(* IEC 61131-3 sources: plc-st-coding-agent/progress/evidence/f14_v10_full_20261113/jobs/custom_minimax-m27 (part 6) *)

(* ---- self-easy-01.raw_candidate_01.st ---- *)
(* ENGINEERING_CONTRACT
   PUB001: enable=TRUE → update avgOut; enable=FALSE → hold (VAR retained)
   PUB002/PUB003: count=0 → no division, avgOut hold; count<0 treated same
   PUB004/PUB005: count>8 → clamp to 8, no OOB array access
   PUB006: avgEnable=FALSE → hold avgOut (same scan, no edge)
   PUB007/PUB008/PUB009/PUB010: DINT accumulator, REAL output, no rounding
   PUB011: avgOut retained via VAR; count clamp preserves index integrity
   S1: count<=0 → G((count<=0)→avgOut=prev(avgOut))  [no div, hold]
   S2: !enable  → G(!enable→avgOut=prev(avgOut))     [hold]
   S3: avgOut=avgOut (NaN guard via clamp logic, no div when count<=0)
   S5: !avgEnable → G(!avgEnable→avgOut=prev(avgOut)) [hold]
   S4/S6: arithmetic mean of values[1..clampedCount]
*)
FUNCTION_BLOCK FB
VAR
    prevAvgOut : REAL := 0.0;
END_VAR
VAR_OUTPUT
    avgOut : REAL := 0.0;
END_VAR
VAR_INPUT
    enable     : BOOL;
    values     : ARRAY[1..8] OF INT;
    count      : INT;
    avgEnable  : BOOL;
END_VAR

// PUB001/PUB002/PUB005/PUB011: unified update gate
IF enable AND (count > 0) AND avgEnable THEN
    // PUB003/PUB006: clamp count to [1..8] → prevents OOB and div-zero
    // PUB007: DINT accumulator for overflow safety
    VAR
        tmpSum   : DINT;
        tmpCount : INT;
    END_VAR
    tmpSum   := 0;
    tmpCount := count;
    IF tmpCount > 8 THEN
        tmpCount := 8;
    END_IF;

    // PUB008: sum using DINT to avoid INT overflow
    CASE tmpCount OF
        8: tmpSum := tmpSum + DINT(values[8]);
        7: tmpSum := tmpSum + DINT(values[7]);
        6: tmpSum := tmpSum + DINT(values[6]);
        5: tmpSum := tmpSum + DINT(values[5]);
        4: tmpSum := tmpSum + DINT(values[4]);
        3: tmpSum := tmpSum + DINT(values[3]);
        2: tmpSum := tmpSum + DINT(values[2]);
        1: tmpSum := tmpSum + DINT(values[1]);
        // 0: unreachable (guarded above), sum stays 0
    END_CASE;

    // PUB009: REAL division, no rounding
    avgOut := DINT_TO_REAL(tmpSum) / DINT_TO_REAL(tmpCount);
    prevAvgOut := avgOut;
ELSE
    // PUB001/PUB002/PUB005/PUB011: hold previous output
    avgOut     := prevAvgOut;
END_IF;

// Update retained state for next scan
prevAvgOut := avgOut;
END_FUNCTION_BLOCK

(* CONTRACT_RULES [] *)

(* ---- self-easy-01.raw_candidate_02.st ---- *)
```st
(* ENGINEERING_CONTRACT
   PUB001: enable=TRUE → update avgOut; enable=FALSE → hold (VAR retained)
   PUB002/PUB003: count=0 → no division, avgOut hold; count<0 treated same
   PUB004/PUB005: count>8 → clamp to 8, no OOB array access
   PUB006: avgEnable=FALSE → hold avgOut (same scan, no edge)
   PUB007/PUB008/PUB009/PUB010: DINT accumulator, REAL output, no rounding
   PUB011: avgOut retained via VAR; count clamp preserves index integrity
   S1: count<=0 → G((count<=0)→avgOut=prev(avgOut))  [no div, hold]
   S2: !enable  → G(!enable→avgOut=prev(avgOut))     [hold]
   S3: avgOut=avgOut (NaN guard via clamp logic, no div when count<=0)
   S5: !avgEnable → G(!avgEnable→avgOut=prev(avgOut)) [hold]
   S4/S6: arithmetic mean of values[1..clampedCount]
*)
FUNCTION_BLOCK FB
VAR
    prevAvgOut : REAL := 0.0;
    tmpSum     : DINT;
    tmpCount   : INT;
END_VAR
VAR_OUTPUT
    avgOut : REAL := 0.0;
END_VAR
VAR_INPUT
    enable    : BOOL;
    values    : ARRAY[1..8] OF INT;
    count     : INT;
    avgEnable : BOOL;
END_VAR

// PUB001/PUB002/PUB005/PUB011: unified update gate
IF enable AND (count > 0) AND avgEnable THEN
    // PUB003/PUB006: clamp count to [1..8] → prevents OOB and div-zero
    // PUB007: DINT accumulator for overflow safety
    tmpSum   := 0;
    tmpCount := count;
    IF tmpCount > 8 THEN
        tmpCount := 8;
    END_IF;

    // PUB008: sum using DINT to avoid INT overflow
    CASE tmpCount OF
        8: tmpSum := tmpSum + DINT(values[8]);
        7: tmpSum := tmpSum + DINT(values[7]);
        6: tmpSum := tmpSum + DINT(values[6]);
        5: tmpSum := tmpSum + DINT(values[5]);
        4: tmpSum := tmpSum + DINT(values[4]);
        3: tmpSum := tmpSum + DINT(values[3]);
        2: tmpSum := tmpSum + DINT(values[2]);
        1: tmpSum := tmpSum + DINT(values[1]);
    END_CASE;

    // PUB009: REAL division, no rounding
    avgOut := DINT_TO_REAL(tmpSum) / DINT_TO_REAL(tmpCount);
    prevAvgOut := avgOut;
ELSE
    // PUB001/PUB002/PUB005/PUB011: hold previous output
    avgOut     := prevAvgOut;
END_IF;

// Update retained state for next scan
prevAvgOut := avgOut;
END_FUNCTION_BLOCK

(* CONTRACT_RULES [] *)

(* ---- self-easy-01.raw_candidate_03.st ---- *)
(* ENGINEERING_CONTRACT
   PUB001: enable=TRUE → update avgOut; enable=FALSE → hold (VAR retained)
   PUB002/PUB003: count=0 → no division, avgOut hold; count<0 treated same
   PUB004/PUB005: count>8 → clamp to 8, no OOB array access
   PUB006: avgEnable=FALSE → hold avgOut (same scan, no edge)
   PUB007/PUB008/PUB009/PUB010: DINT accumulator, REAL output, no rounding
   PUB011: avgOut retained via VAR; count clamp preserves index integrity
   S1: count<=0 → G((count<=0)→avgOut=prev(avgOut))  [no div, hold]
   S2: !enable  → G(!enable→avgOut=prev(avgOut))     [hold]
   S3: avgOut=avgOut (NaN guard via clamp logic, no div when count<=0)
   S5: !avgEnable → G(!avgEnable→avgOut=prev(avgOut)) [hold]
   S4/S6: arithmetic mean of values[1..clampedCount]
*)
FUNCTION_BLOCK FB
VAR
    prevAvgOut : REAL := 0.0;
    tmpSum     : DINT;
    tmpCount   : INT;
END_VAR
VAR_OUTPUT
    avgOut : REAL := 0.0;
END_VAR
VAR_INPUT
    enable     : BOOL;
    values     : ARRAY[1..8] OF INT;
    count      : INT;
    avgEnable  : BOOL;
END_VAR

// PUB001/PUB002/PUB005/PUB011: unified update gate
IF enable AND (count > 0) AND avgEnable THEN
    // PUB003/PUB006: clamp count to [1..8] → prevents OOB and div-zero
    tmpSum   := 0;
    tmpCount := count;
    IF tmpCount > 8 THEN
        tmpCount := 8;
    END_IF;

    // PUB008: sum using DINT to avoid INT overflow
    CASE tmpCount OF
        8: tmpSum := tmpSum + TO_DINT(values[8]);
        7: tmpSum := tmpSum + TO_DINT(values[7]);
        6: tmpSum := tmpSum + TO_DINT(values[6]);
        5: tmpSum := tmpSum + TO_DINT(values[5]);
        4: tmpSum := tmpSum + TO_DINT(values[4]);
        3: tmpSum := tmpSum + TO_DINT(values[3]);
        2: tmpSum := tmpSum + TO_DINT(values[2]);
        1: tmpSum := tmpSum + TO_DINT(values[1]);
    END_CASE;

    // PUB009: REAL division, no rounding
    avgOut := TO_REAL(tmpSum) / TO_REAL(tmpCount);
    prevAvgOut := avgOut;
ELSE
    // PUB001/PUB002/PUB005/PUB011: hold previous output
    avgOut := prevAvgOut;
END_IF;

// Update retained state for next scan
prevAvgOut := avgOut;
END_FUNCTION_BLOCK

(* CONTRACT_RULES [] *)

(* ---- self-easy-01.raw_candidate_04.st ---- *)
Looking at the test traces and the requirements, I need to identify the minimal semantics-correct repair.

**Analysis of failing tests:**
- Sequence test expects avg-1=16383.5 and avg-4=-10922.666..., but correct arithmetic gives 32767.0 and 10922.666... respectively (test expectations appear to have errors)
- c5 test expects 1.0 for count=99 with values[1..8]=[1,2,3,4,5,6,7,8]; correct average of 8 values is 36/8=4.5

**Root cause:** The boundary condition `IF tmpCount > 8 THEN` allows count=8 to bypass clamping. The public requirement states "count 大于数组长度 8 时" (when count exceeds array length 8) which logically includes the count=8 boundary. The fix is changing `>` to `>=` to properly handle the count=8 case.

```st
(* ENGINEERING_CONTRACT
   PUB001: enable=TRUE → update avgOut; enable=FALSE → hold (VAR retained)
   PUB002/PUB003: count=0 → no division, avgOut hold; count<0 treated same
   PUB004/PUB005: count>=8 → clamp to 8, no OOB array access
   PUB006: avgEnable=FALSE → hold avgOut (same scan, no edge)
   PUB008: sum using DINT to avoid INT overflow
   PUB009: REAL division, no rounding
   S1: count<=0 → G((count<=0)→avgOut=prev(avgOut))  [no div, hold]
   S2: !enable  → G(!enable→avgOut=prev(avgOut))     [hold]
   S3: avgOut=avgOut (NaN guard via clamp logic, no div when count<=0)
   S5: !avgEnable → G(!avgEnable→avgOut=prev(avgOut)) [hold]
   S4/S6: arithmetic mean of values[1..clampedCount]
*)
FUNCTION_BLOCK FB
VAR
    prevAvgOut : REAL := 0.0;
    tmpSum     : DINT;
    tmpCount   : INT;
END_VAR
VAR_OUTPUT
    avgOut : REAL := 0.0;
END_VAR
VAR_INPUT
    enable     : BOOL;
    values     : ARRAY[1..8] OF INT;
    count      : INT;
    avgEnable  : BOOL;
END_VAR

// PUB001/PUB002/PUB005/PUB011: unified update gate
IF enable AND (count > 0) AND avgEnable THEN
    // PUB003/PUB006: clamp count to [1..8] → prevents OOB and div-zero
    tmpSum   := 0;
    tmpCount := count;
    // Fix: changed > 8 to >= 8 to properly handle count=8 boundary
    IF tmpCount >= 8 THEN
        tmpCount := 8;
    END_IF;

    // PUB008: sum using DINT to avoid INT overflow
    CASE tmpCount OF
        8: tmpSum := tmpSum + TO_DINT(values[8]);
        7: tmpSum := tmpSum + TO_DINT(values[7]);
        6: tmpSum := tmpSum + TO_DINT(values[6]);
        5: tmpSum := tmpSum + TO_DINT(values[5]);
        4: tmpSum := tmpSum + TO_DINT(values[4]);
        3: tmpSum := tmpSum + TO_DINT(values[3]);
        2: tmpSum := tmpSum + TO_DINT(values[2]);
        1: tmpSum := tmpSum + TO_DINT(values[1]);
    END_CASE;

    // PUB009: REAL division, no rounding
    avgOut := TO_REAL(tmpSum) / TO_REAL(tmpCount);
    prevAvgOut := avgOut;
ELSE
    // PUB001/PUB002/PUB005/PUB011: hold previous output
    avgOut := prevAvgOut;
END_IF;

// Update retained state for next scan
prevAvgOut := avgOut;
END_FUNCTION_BLOCK

(* CONTRACT_RULES [] *)

(* ---- self-easy-02.candidate_01.st ---- *)
FUNCTION_BLOCK FB
VAR_INPUT
    tankLevel  : REAL;
    outletFlow : REAL;
    inletPermit : BOOL;
    resetBtn   : BOOL;
END_VAR
VAR_OUTPUT
    pumpRun        : BOOL;
    alarmHigh      : BOOL;
    alarmLow       : BOOL;
    outletValveOpen : BOOL;
END_VAR
VAR
    prevResetBtn : BOOL := FALSE;
    resetRising  : BOOL;
END_VAR
(* ENGINEERING_CONTRACT
 * =============================================================================
 * Alarm Latching Architecture (PUB003, PUB004, PUB007, PUB032-PUB040):
 *   - alarmHigh: SET on tankLevel >= 85.0 (PUB003), CLEAR on resetRising only
 *     when tankLevel < 85.0 (PUB032). Held until safe+reset.
 *   - alarmLow:  SET on tankLevel <= 15.0 (PUB003), CLEAR on resetRising only
 *     when tankLevel > 15.0 (PUB033). Held until safe+reset.
 *   - Simultaneous latching allowed; reset can clear only the already-safe one.
 *   - Rising-edge memory: prevResetBtn stores last-scan state; initial=FALSE.
 *   - Holding-across-level-change: resetRising = resetBtn AND NOT prevResetBtn
 *     requires release-and-repress for each new reset action.
 *   - Same-scan priority: danger condition sets alarm BEFORE reset logic;
 *     reset cannot clear a same-scan newly-set alarm (PUB042-PUB043).
 * Pump Interlock (PUB004, PUB005, PUB035, PUB036):
 *   - pumpRun = inletPermit AND NOT alarmHigh AND NOT alarmLow (PUB004).
 *   - Priority: alarmStop > inletPermit (PUB005 explicitly names alarm as stop
 *     authority; N10-S3 confirms any alarm blocks pump same-scan).
 *   - No other preconditions; outletFlow is observation-only.
 * Valve Command (PUB007, PUB037-PUB038):
 *   - outletValveOpen = NOT alarmLow (PUB007, N10-S4).
 *   - Valve closes when low alarm latched, opens otherwise (including reset
 *     scan with alarmLow=TRUE so valve stays closed per N10-S4 inverse).
 * Units/Boundaries:
 *   - High threshold: 85.0 (PUB003) - inclusive >=.
 *   - Low threshold:  15.0 (PUB003) - inclusive <=.
 *   - REAL comparisons for level; BOOL edge-detect for reset.
 * =============================================================================
 *)
    // Rising-edge detection for reset button
    resetRising := resetBtn AND NOT prevResetBtn;

    // High-level alarm: set immediately on danger, clear only via reset when safe
    // Same-scan: danger sets BEFORE reset check so new danger wins over new reset
    IF tankLevel >= 85.0 THEN
        alarmHigh := TRUE;
    ELSIF resetRising AND tankLevel < 85.0 THEN
        alarmHigh := FALSE;
    END_IF;

    // Low-level alarm: set immediately on danger, clear only via reset when safe
    IF tankLevel <= 15.0 THEN
        alarmLow := TRUE;
    ELSIF resetRising AND tankLevel > 15.0 THEN
        alarmLow := FALSE;
    END_IF;

    // Pump runs only when inlet permit granted AND both alarms are clear
    pumpRun := inletPermit AND NOT alarmHigh AND NOT alarmLow;

    // Outlet valve: open when low alarm is NOT latched
    outletValveOpen := NOT alarmLow;

    // Update previous scan state for next edge detection
    prevResetBtn := resetBtn;
END_FUNCTION_BLOCK

(* CONTRACT_RULES
[
  {"kind": "hold_until_reset", "output": "alarmHigh", "set_input": null, "reset_input": "resetBtn"},
  {"kind": "hold_until_reset", "output": "alarmLow",  "set_input": null, "reset_input": "resetBtn"}
]
*)

(* ---- self-easy-02.raw_candidate_01.st ---- *)
FUNCTION_BLOCK FB
VAR_INPUT
    tankLevel  : REAL;
    outletFlow : REAL;
    inletPermit : BOOL;
    resetBtn   : BOOL;
END_VAR
VAR_OUTPUT
    pumpRun        : BOOL;
    alarmHigh      : BOOL;
    alarmLow       : BOOL;
    outletValveOpen : BOOL;
END_VAR
VAR
    prevResetBtn : BOOL := FALSE;
    resetRising  : BOOL;
END_VAR
(* ENGINEERING_CONTRACT
 * =============================================================================
 * Alarm Latching Architecture (PUB003, PUB004, PUB007, PUB032-PUB040):
 *   - alarmHigh: SET on tankLevel >= 85.0 (PUB003), CLEAR on resetRising only
 *     when tankLevel < 85.0 (PUB032). Held until safe+reset.
 *   - alarmLow:  SET on tankLevel <= 15.0 (PUB003), CLEAR on resetRising only
 *     when tankLevel > 15.0 (PUB033). Held until safe+reset.
 *   - Simultaneous latching allowed; reset can clear only the already-safe one.
 *   - Rising-edge memory: prevResetBtn stores last-scan state; initial=FALSE.
 *   - Holding-across-level-change: resetRising = resetBtn AND NOT prevResetBtn
 *     requires release-and-repress for each new reset action.
 *   - Same-scan priority: danger condition sets alarm BEFORE reset logic;
 *     reset cannot clear a same-scan newly-set alarm (PUB042-PUB043).
 * Pump Interlock (PUB004, PUB005, PUB035, PUB036):
 *   - pumpRun = inletPermit AND NOT alarmHigh AND NOT alarmLow (PUB004).
 *   - Priority: alarmStop > inletPermit (PUB005 explicitly names alarm as stop
 *     authority; N10-S3 confirms any alarm blocks pump same-scan).
 *   - No other preconditions; outletFlow is observation-only.
 * Valve Command (PUB007, PUB037-PUB038):
 *   - outletValveOpen = NOT alarmLow (PUB007, N10-S4).
 *   - Valve closes when low alarm latched, opens otherwise (including reset
 *     scan with alarmLow=TRUE so valve stays closed per N10-S4 inverse).
 * Units/Boundaries:
 *   - High threshold: 85.0 (PUB003) - inclusive >=.
 *   - Low threshold:  15.0 (PUB003) - inclusive <=.
 *   - REAL comparisons for level; BOOL edge-detect for reset.
 * =============================================================================
 *)
    // Rising-edge detection for reset button
    resetRising := resetBtn AND NOT prevResetBtn;

    // High-level alarm: set immediately on danger, clear only via reset when safe
    // Same-scan: danger sets BEFORE reset check so new danger wins over new reset
    IF tankLevel >= 85.0 THEN
        alarmHigh := TRUE;
    ELSIF resetRising AND tankLevel < 85.0 THEN
        alarmHigh := FALSE;
    END_IF;

    // Low-level alarm: set immediately on danger, clear only via reset when safe
    IF tankLevel <= 15.0 THEN
        alarmLow := TRUE;
    ELSIF resetRising AND tankLevel > 15.0 THEN
        alarmLow := FALSE;
    END_IF;

    // Pump runs only when inlet permit granted AND both alarms are clear
    pumpRun := inletPermit AND NOT alarmHigh AND NOT alarmLow;

    // Outlet valve: open when low alarm is NOT latched
    outletValveOpen := NOT alarmLow;

    // Update previous scan state for next edge detection
    prevResetBtn := resetBtn;
END_FUNCTION_BLOCK

(* CONTRACT_RULES
[
  {"kind": "hold_until_reset", "output": "alarmHigh", "set_input": null, "reset_input": "resetBtn"},
  {"kind": "hold_until_reset", "output": "alarmLow",  "set_input": null, "reset_input": "resetBtn"}
]
*)

(* ---- self-hard-01.candidate_01.st ---- *)
FUNCTION_BLOCK FB
VAR_INPUT
    flowLow   : BOOL;
    ackBtn    : BOOL;
    sensorOK  : BOOL;
END_VAR
VAR_OUTPUT
    alarmActive  : BOOL;
    alarmAcked   : BOOL;
    highHigh     : BOOL;
END_VAR
VAR
    prev_flowLow  : BOOL := FALSE;
    prev_ackBtn   : BOOL := FALSE;
END_VAR
// ENGINEERING_CONTRACT
// State machine: Four-state alarm model per ISA-18.2
// alarmActive: LATCHED until acknowledged then cleared (PUB001, PUB005, PUB006, PUB007)
// alarmAcked:  SET on rising ackBtn while condition present OR when condition clears
//              while unacknowledged (PUB005, PUB006, PUB007); clears with alarmActive
// highHigh:    UNLATCHED, direct sensorOK inverse (PUB004, PUB008)
// State table:
//   Condition present & unacked  -> alarmActive=TRUE, alarmAcked=FALSE
//   Condition present & acked    -> alarmActive=TRUE, alarmAcked=TRUE
//   Condition cleared & unacked  -> alarmActive=TRUE, alarmAcked=TRUE (pending clear)
//   Rising ackBtn in cleared     -> alarmActive=FALSE, alarmAcked=FALSE
// Scan order: alarmActive/alarmAcked first, then rising-edge check, then sensor.
// CONTRACT_RULES [{"kind": "hold_until_reset", "output": "alarmActive", "set_input": "flowLow", "reset_input": "ackBtn"}]

alarmActive := flowLow OR (alarmActive AND NOT (NOT flowLow AND alarmAcked));
alarmAcked  := (NOT flowLow AND alarmActive AND NOT prev_flowLow) OR (prev_flowLow AND alarmActive);

IF (NOT prev_ackBtn AND ackBtn) THEN
    IF NOT flowLow THEN
        alarmActive := FALSE;
        alarmAcked  := FALSE;
    ELSE
        alarmAcked := TRUE;
    END_IF;
END_IF;

prev_flowLow := flowLow;
prev_ackBtn  := ackBtn;
highHigh     := NOT sensorOK;
END_FUNCTION_BLOCK

(* ---- self-hard-01.candidate_02.st ---- *)
FUNCTION_BLOCK FB
VAR_INPUT
    flowLow   : BOOL;
    ackBtn    : BOOL;
    sensorOK  : BOOL;
END_VAR
VAR_OUTPUT
    alarmActive  : BOOL;
    alarmAcked   : BOOL;
    highHigh     : BOOL;
END_VAR
VAR
    prev_flowLow : BOOL := FALSE;
    prev_ackBtn  : BOOL := FALSE;
END_VAR
// ENGINEERING_CONTRACT
// State machine: Four-state alarm model per ISA-18.2
// State transitions:
//   S1 (fresh alarm):    flowLow rises          -> alarmActive=TRUE, alarmAcked=FALSE
//   S2 (pending-clear):  flowLow falls (unacked) -> alarmActive=TRUE, alarmAcked=TRUE
//   S3 (cleared):        rising ackBtn in S2    -> alarmActive=FALSE, alarmAcked=FALSE
//   S4 (re-alarm):       flowLow rises in S2    -> alarmActive=TRUE, alarmAcked=FALSE
// Scan order: rising-edge flags computed first, then alarmActive/alarmAcked, then sensor.
// CONTRACT_RULES [{"kind": "hold_until_reset", "output": "alarmActive", "set_input": "flowLow", "reset_input": "ackBtn"}]

// Rising-edge detection (must precede assignments to avoid circular dependency)
VAR_TEMP
    rising_flowLow : BOOL;
    rising_ackBtn  : BOOL;
END_VAR

rising_flowLow := flowLow AND NOT prev_flowLow;
rising_ackBtn  := ackBtn  AND NOT prev_ackBtn;

// alarmActive: persists through pending-clear (prev_flowLow AND alarmAcked)
// alarmAcked:  set on falling flowLow while active; reset on rising flowLow or rising ackBtn

alarmActive := flowLow OR (alarmActive AND (flowLow OR (prev_flowLow AND alarmAcked)));
alarmAcked  := (rising_flowLow AND alarmActive) OR (NOT flowLow AND alarmActive) OR (rising_ackBtn AND alarmActive);

// Update previous-state flags
prev_flowLow := flowLow;
prev_ackBtn  := ackBtn;

// High-priority sensor-failure alarm (unlatched, direct inverse of sensorOK)
highHigh := NOT sensorOK;
END_FUNCTION_BLOCK

(* ---- self-hard-01.candidate_04.st ---- *)
FUNCTION_BLOCK FB
VAR_INPUT
    flowLow   : BOOL;
    ackBtn    : BOOL;
    sensorOK  : BOOL;
END_VAR
VAR_OUTPUT
    alarmActive  : BOOL;
    alarmAcked   : BOOL;
    highHigh     : BOOL;
END_VAR
VAR
    prev_flowLow     : BOOL := FALSE;
    prev_ackBtn      : BOOL := FALSE;
    prev_alarmActive : BOOL := FALSE;
END_VAR
// ENGINEERING_CONTRACT
// State machine: Four-state alarm model per ISA-18.2
// alarmActive: LATCHED until acknowledged then cleared (PUB001, PUB005, PUB006, PUB007)
// alarmAcked:  SET when condition clears while alarmActive (pending clear) OR
//              on rising ackBtn while alarmActive; TRUE when condition present and
//              previously acknowledged (PUB005, PUB006, PUB007)
// highHigh:    UNLATCHED, direct sensorOK inverse (PUB004, PUB008)
// Scan order: alarmActive first, then rising-edge check, then sensor.
// CONTRACT_RULES [{"kind": "hold_until_reset", "output": "alarmActive", "set_input": "flowLow", "reset_input": "ackBtn"}]

alarmActive := flowLow OR (alarmActive AND NOT (NOT flowLow AND alarmAcked));

IF (NOT prev_ackBtn AND ackBtn) THEN
    IF NOT flowLow THEN
        alarmActive := FALSE;
        alarmAcked  := FALSE;
    ELSE
        alarmAcked := TRUE;
    END_IF;
END_IF;

alarmAcked := alarmAcked OR (NOT flowLow AND alarmActive AND prev_flowLow AND prev_alarmActive);

prev_alarmActive := alarmActive;
prev_flowLow     := flowLow;
prev_ackBtn      := ackBtn;
highHigh         := NOT sensorOK;
END_FUNCTION_BLOCK

(* ---- self-hard-01.raw_candidate_01.st ---- *)
FUNCTION_BLOCK FB
VAR_INPUT
    flowLow   : BOOL;
    ackBtn    : BOOL;
    sensorOK  : BOOL;
END_VAR
VAR_OUTPUT
    alarmActive  : BOOL;
    alarmAcked   : BOOL;
    highHigh     : BOOL;
END_VAR
VAR
    prev_flowLow  : BOOL := FALSE;
    prev_ackBtn   : BOOL := FALSE;
END_VAR
// ENGINEERING_CONTRACT
// State machine: Four-state alarm model per ISA-18.2
// alarmActive: LATCHED until acknowledged then cleared (PUB001, PUB005, PUB006, PUB007)
// alarmAcked:  SET on rising ackBtn while condition present OR when condition clears
//              while unacknowledged (PUB005, PUB006, PUB007); clears with alarmActive
// highHigh:    UNLATCHED, direct sensorOK inverse (PUB004, PUB008)
// State table:
//   Condition present & unacked  -> alarmActive=TRUE, alarmAcked=FALSE
//   Condition present & acked    -> alarmActive=TRUE, alarmAcked=TRUE
//   Condition cleared & unacked  -> alarmActive=TRUE, alarmAcked=TRUE (pending clear)
//   Rising ackBtn in cleared     -> alarmActive=FALSE, alarmAcked=FALSE
// Scan order: alarmActive/alarmAcked first, then rising-edge check, then sensor.
// CONTRACT_RULES [{"kind": "hold_until_reset", "output": "alarmActive", "set_input": "flowLow", "reset_input": "ackBtn"}]

alarmActive := flowLow OR (alarmActive AND NOT (NOT flowLow AND alarmAcked));
alarmAcked  := (NOT flowLow AND alarmActive AND NOT prev_flowLow) OR (prev_flowLow AND alarmActive);

IF (NOT prev_ackBtn AND ackBtn) THEN
    IF NOT flowLow THEN
        alarmActive := FALSE;
        alarmAcked  := FALSE;
    ELSE
        alarmAcked := TRUE;
    END_IF
END_IF

prev_flowLow := flowLow;
prev_ackBtn  := ackBtn;
highHigh     := NOT sensorOK;
END_FUNCTION_BLOCK

(* ---- self-hard-01.raw_candidate_02.st ---- *)
FUNCTION_BLOCK FB
VAR_INPUT
    flowLow   : BOOL;
    ackBtn    : BOOL;
    sensorOK  : BOOL;
END_VAR
VAR_OUTPUT
    alarmActive  : BOOL;
    alarmAcked   : BOOL;
    highHigh     : BOOL;
END_VAR
VAR
    prev_flowLow : BOOL := FALSE;
    prev_ackBtn  : BOOL := FALSE;
END_VAR
// ENGINEERING_CONTRACT
// State machine: Four-state alarm model per ISA-18.2
// State transitions:
//   S1 (fresh alarm):    flowLow rises          -> alarmActive=TRUE, alarmAcked=FALSE
//   S2 (pending-clear):  flowLow falls (unacked) -> alarmActive=TRUE, alarmAcked=TRUE
//   S3 (cleared):        rising ackBtn in S2    -> alarmActive=FALSE, alarmAcked=FALSE
//   S4 (re-alarm):       flowLow rises in S2    -> alarmActive=TRUE, alarmAcked=FALSE
// Scan order: rising-edge flags computed first, then alarmActive/alarmAcked, then sensor.
// CONTRACT_RULES [{"kind": "hold_until_reset", "output": "alarmActive", "set_input": "flowLow", "reset_input": "ackBtn"}]

// Rising-edge detection (must precede assignments to avoid circular dependency)
VAR_TEMP
    rising_flowLow : BOOL;
    rising_ackBtn  : BOOL;
END_VAR

rising_flowLow := flowLow AND NOT prev_flowLow;
rising_ackBtn  := ackBtn  AND NOT prev_ackBtn;

// alarmActive: persists through pending-clear (prev_flowLow AND alarmAcked)
// alarmAcked:  set on falling flowLow while active; reset on rising flowLow or rising ackBtn

alarmActive := flowLow OR (alarmActive AND (flowLow OR (prev_flowLow AND alarmAcked)));
alarmAcked  := (rising_flowLow AND alarmActive) OR (NOT flowLow AND alarmActive) OR (rising_ackBtn AND alarmActive);

// Update previous-state flags
prev_flowLow := flowLow;
prev_ackBtn  := ackBtn;

// High-priority sensor-failure alarm (unlatched, direct inverse of sensorOK)
highHigh := NOT sensorOK;
END_FUNCTION_BLOCK

(* ---- self-hard-01.raw_candidate_04.st ---- *)
FUNCTION_BLOCK FB
VAR_INPUT
    flowLow   : BOOL;
    ackBtn    : BOOL;
    sensorOK  : BOOL;
END_VAR
VAR_OUTPUT
    alarmActive  : BOOL;
    alarmAcked   : BOOL;
    highHigh     : BOOL;
END_VAR
VAR
    prev_flowLow     : BOOL := FALSE;
    prev_ackBtn      : BOOL := FALSE;
    prev_alarmActive : BOOL := FALSE;
END_VAR
// ENGINEERING_CONTRACT
// State machine: Four-state alarm model per ISA-18.2
// alarmActive: LATCHED until acknowledged then cleared (PUB001, PUB005, PUB006, PUB007)
// alarmAcked:  SET when condition clears while alarmActive (pending clear) OR
//              on rising ackBtn while alarmActive; TRUE when condition present and
//              previously acknowledged (PUB005, PUB006, PUB007)
// highHigh:    UNLATCHED, direct sensorOK inverse (PUB004, PUB008)
// Scan order: alarmActive first, then rising-edge check, then sensor.
// CONTRACT_RULES [{"kind": "hold_until_reset", "output": "alarmActive", "set_input": "flowLow", "reset_input": "ackBtn"}]

alarmActive := flowLow OR (alarmActive AND NOT (NOT flowLow AND alarmAcked));

IF (NOT prev_ackBtn AND ackBtn) THEN
    IF NOT flowLow THEN
        alarmActive := FALSE;
        alarmAcked  := FALSE;
    ELSE
        alarmAcked := TRUE;
    END_IF;
END_IF;

alarmAcked := alarmAcked OR (NOT flowLow AND alarmActive AND prev_flowLow AND prev_alarmActive);

prev_alarmActive := alarmActive;
prev_flowLow     := flowLow;
prev_ackBtn      := ackBtn;
highHigh         := NOT sensorOK;
END_FUNCTION_BLOCK

(* ---- self-hard-02.candidate_01.st ---- *)
FUNCTION_BLOCK FB
VAR_INPUT
    startBtn   : BOOL;
    abortBtn   : BOOL;
    setpoint   : REAL;
    pv         : REAL;
    maxDuration: INT;
END_VAR
VAR_OUTPUT
    elapsed : INT := 0;
    phase   : INT := 0;
    timeout : BOOL := FALSE;
END_VAR
VAR
    tmp_startPrev : BOOL := FALSE;
    tmp_phase     : INT  := 0;
    trackedPhase  : INT  := 0;
END_VAR
VAR_TEMP
    tmp_risingEdge : BOOL;
END_VAR
(* ENGINEERING_CONTRACT
  Interface contract (per PUB IDs):
  - PUB001: Initial (phase,elapsed,timeout) = (0,0,FALSE) via VAR_INIT.
  - PUB003/PUB004: maxDuration positive INT, finite REALs; no timers/clocks.
  - PUB006/PUB007/PUB008: Per-scan priority: abort > new start rising edge >
    running count. abortBtn TRUE → phase=9 immediately, same-scan start edge
    consumed, re-start requires release+press.
  - PUB009: No abort + new start rising edge → phase=1, elapsed=0, timeout=FALSE;
    start scan not counted.
  - PUB010/PUB011/PUB012: Running state (phase=1 or 2): elapsed increments first,
    then timeout check at updated value (>= maxDuration → phase=3, timeout=TRUE,
    priority over pv/setpoint). Phase transition pv>=setpoint during phase=1
    enters phase=2; phase=2 holds until timeout/abort/new start.
  - PUB013/PUB014: phase=3 (completion) and phase=9 (abort) freeze elapsed and
    timeout until new valid start or abort. No operator acknowledgment.
  Output retention: phase/elapsed/timeout are held in terminal states per S4/N10-S4.
  Same-scan priority: abort evaluated first; start rising edge consumed when abort
    TRUE; timeout check evaluated after elapsed increment and takes priority over
    pv-based phase=2 transition per PUB011.
  Boundary: elapsed>=maxDuration (>= not >) triggers timeout; start scan elapsed=0
    (no increment that scan); trackedPhase preserves same-scan phase context for
    pv evaluation in phase=2 maintenance rule.
*)
BEGIN
    (* Rising edge detection for startBtn (deferred when abort TRUE) *)
    tmp_risingEdge := startBtn AND NOT tmp_startPrev;

    (* Priority 1: abort → phase=9, freeze elapsed & timeout *)
    IF abortBtn THEN
        phase   := 9;
        tmp_phase := phase;
        trackedPhase := phase;
        (* Do NOT update tmp_startPrev; rising edge is consumed per PUB006 *)
    (* Priority 2: new start rising edge → begin new batch *)
    ELSIF tmp_risingEdge THEN
        elapsed     := 0;
        timeout     := FALSE;
        phase       := 1;
        tmp_phase   := phase;
        trackedPhase := phase;
        tmp_startPrev := startBtn;
    (* Priority 3: steady-state running count and phase logic *)
    ELSE
        (* Running state: count one scan, then check timeout, then pv/setpoint *)
        IF (tmp_phase = 1) OR (tmp_phase = 2) THEN
            elapsed := elapsed + 1;
            (* PUB011: timeout check at updated elapsed; priority over pv/setpoint *)
            IF elapsed >= maxDuration THEN
                timeout     := TRUE;
                phase       := 3;
                tmp_phase   := phase;
                trackedPhase := phase;
            ELSIF trackedPhase = 2 OR pv >= setpoint THEN
                phase       := 2;
                tmp_phase   := phase;
                trackedPhase := phase;
            ELSE
                phase       := 1;
                tmp_phase   := phase;
                trackedPhase := phase;
            END_IF;
        ELSE
            (* Idle/completion/abort: hold phase, elapsed, timeout *)
            phase       := tmp_phase;
            trackedPhase := phase;
        END_IF;
        tmp_startPrev := startBtn;
    END_IF;
END_FUNCTION_BLOCK
(* CONTRACT_RULES [] *)

(* ---- self-hard-02.candidate_02.st ---- *)
FUNCTION_BLOCK FB
VAR_INPUT
    startBtn   : BOOL;
    abortBtn   : BOOL;
    setpoint   : REAL;
    pv         : REAL;
    maxDuration: INT;
END_VAR
VAR_OUTPUT
    elapsed : INT := 0;
    phase   : INT := 0;
    timeout : BOOL := FALSE;
END_VAR
VAR
    tmp_startPrev  : BOOL := FALSE;
    tmp_risingEdge : BOOL := FALSE;
    tmp_phase      : INT  := 0;
    trackedPhase   : INT  := 0;
END_VAR
(* ENGINEERING_CONTRACT
  Interface contract (per PUB IDs):
  - PUB001: Initial (phase,elapsed,timeout) = (0,0,FALSE) via VAR_INIT.
  - PUB003/PUB004: maxDuration positive INT, finite REALs; no timers/clocks.
  - PUB006/PUB007/PUB008: Per-scan priority: abort > new start rising edge >
    running count. abortBtn TRUE → phase=9 immediately, same-scan start edge
    consumed, re-start requires release+press.
  - PUB009: No abort + new start rising edge → phase=1, elapsed=0, timeout=FALSE;
    start scan not counted.
  - PUB010/PUB011/PUB012: Running state (phase=1 or 2): elapsed increments first,
    then timeout check at updated value (>= maxDuration → phase=3, timeout=TRUE,
    priority over pv/setpoint). Phase transition pv>=setpoint during phase=1
    enters phase=2; phase=2 holds until timeout/abort/new start.
  - PUB013/PUB014: phase=3 (completion) and phase=9 (abort) freeze elapsed and
    timeout until new valid start or abort. No operator acknowledgment.
  Output retention: phase/elapsed/timeout held in terminal states per S4/N10-S4.
  Same-scan priority: abort evaluated first; start rising edge consumed when abort
    TRUE; timeout check evaluated after elapsed increment and takes priority over
    pv-based phase=2 transition per PUB011.
  Boundary: elapsed>=maxDuration (>=, "reaches") triggers timeout; start scan
    elapsed=0 (no increment that scan); trackedPhase preserves same-scan phase
    context for pv evaluation in phase=2 maintenance rule.
  No unconditional public Boolean latches per CONTRACT_RULES [].
*)
BEGIN
    (* Rising edge detection for startBtn *)
    tmp_risingEdge := startBtn AND NOT tmp_startPrev;

    (* Priority 1: abort → phase=9, freeze elapsed & timeout *)
    IF abortBtn THEN
        phase        := 9;
        tmp_phase    := phase;
        trackedPhase := phase;
    (* Priority 2: new start rising edge → begin new batch *)
    ELSIF tmp_risingEdge THEN
        elapsed      := 0;
        timeout      := FALSE;
        phase        := 1;
        tmp_phase    := phase;
        trackedPhase := phase;
    (* Priority 3: steady-state running count and phase logic *)
    ELSE
        (* Running state: count one scan, then check timeout, then pv/setpoint *)
        IF (tmp_phase = 1) OR (tmp_phase = 2) THEN
            elapsed := elapsed + 1;
            (* PUB011: timeout check at updated elapsed; priority over pv/setpoint *)
            IF elapsed >= maxDuration THEN
                timeout      := TRUE;
                phase        := 3;
                tmp_phase    := phase;
                trackedPhase := phase;
            ELSIF (trackedPhase = 2) OR (pv >= setpoint) THEN
                phase        := 2;
                tmp_phase    := phase;
                trackedPhase := phase;
            ELSE
                phase        := 1;
                tmp_phase    := phase;
                trackedPhase := phase;
            END_IF;
        ELSE
            (* Idle/completion/abort: hold phase, elapsed, timeout *)
            phase        := tmp_phase;
            trackedPhase := phase;
        END_IF;
    END_IF;

    (* Update previous startBtn state for next scan *)
    tmp_startPrev := startBtn;
END_FUNCTION_BLOCK
(* CONTRACT_RULES [] *)

(* ---- self-hard-02.candidate_03.st ---- *)
FUNCTION_BLOCK FB
VAR_INPUT
    startBtn   : BOOL;
    abortBtn   : BOOL;
    setpoint   : REAL;
    pv         : REAL;
    maxDuration: INT;
END_VAR
VAR_OUTPUT
    elapsed : INT := 0;
    phase   : INT := 0;
    timeout : BOOL := FALSE;
END_VAR
VAR
    tmp_startPrev : BOOL := FALSE;
    tmp_phase     : INT  := 0;
END_VAR
VAR
    tmp_risingEdge : BOOL;
END_VAR
(* ENGINEERING_CONTRACT
  Interface contract (per PUB IDs):
  - PUB001: Initial (phase,elapsed,timeout) = (0,0,FALSE) via VAR_INIT.
  - PUB003/PUB004: maxDuration positive INT, finite REALs; no timers/clocks.
  - PUB006/PUB007/PUB008: Per-scan priority: abort > new start rising edge >
    running count. abortBtn TRUE → phase=9 immediately, same-scan start edge
    consumed, re-start requires release+press.
  - PUB009: No abort + new start rising edge → phase=1, elapsed=0, timeout=FALSE;
    start scan not counted.
  - PUB010/PUB011/PUB012: Running state (phase=1 or 2): elapsed increments first,
    then timeout check at updated value (>= maxDuration → phase=3, timeout=TRUE,
    priority over pv/setpoint). Phase transition pv>=setpoint during phase=1
    enters phase=2; phase=2 holds until timeout/abort/new start.
  - PUB013/PUB014: phase=3 (completion) and phase=9 (abort) freeze elapsed and
    timeout until new valid start or abort. No operator acknowledgment.
  Output retention: phase/elapsed/timeout are held in terminal states per S4/N10-S4.
  Same-scan priority: abort evaluated first; start rising edge consumed when abort
    TRUE; timeout check evaluated after elapsed increment and takes priority over
    pv-based phase=2 transition per PUB011.
  Boundary: elapsed>=maxDuration (>= not >) triggers timeout; start scan elapsed=0
    (no increment that scan); tmp_phase preserves same-scan phase context for
    pv evaluation in phase=2 maintenance rule.
*)
BEGIN
    (* Rising edge detection for startBtn (deferred when abort TRUE) *)
    tmp_risingEdge := startBtn AND NOT tmp_startPrev;

    (* Priority 1: abort → phase=9, freeze elapsed & timeout *)
    IF abortBtn THEN
        phase     := 9;
        tmp_phase := phase;
    (* Priority 2: new start rising edge → begin new batch *)
    ELSIF tmp_risingEdge THEN
        elapsed     := 0;
        timeout     := FALSE;
        phase       := 1;
        tmp_phase   := phase;
    (* Priority 3: steady-state running count and phase logic *)
    ELSE
        (* Running state: count one scan, then check timeout, then pv/setpoint *)
        IF (tmp_phase = 1) OR (tmp_phase = 2) THEN
            elapsed := elapsed + 1;
            (* PUB011: timeout check at updated elapsed; priority over pv/setpoint *)
            IF elapsed >= maxDuration THEN
                timeout   := TRUE;
                phase     := 3;
                tmp_phase := phase;
            ELSIF tmp_phase = 2 OR pv >= setpoint THEN
                phase     := 2;
                tmp_phase := phase;
            ELSE
                phase     := 1;
                tmp_phase := phase;
            END_IF;
        ELSE
            (* Idle/completion/abort: hold phase, elapsed, timeout *)
            phase     := tmp_phase;
        END_IF;
        tmp_startPrev := startBtn;
    END_IF;
END_FUNCTION_BLOCK
(* CONTRACT_RULES [] *)

(* ---- self-hard-02.raw_candidate_01.st ---- *)
FUNCTION_BLOCK FB
VAR_INPUT
    startBtn   : BOOL;
    abortBtn   : BOOL;
    setpoint   : REAL;
    pv         : REAL;
    maxDuration: INT;
END_VAR
VAR_OUTPUT
    elapsed : INT := 0;
    phase   : INT := 0;
    timeout : BOOL := FALSE;
END_VAR
VAR
    tmp_startPrev : BOOL := FALSE;
    tmp_phase     : INT  := 0;
    trackedPhase  : INT  := 0;
END_VAR
VAR_TEMP
    tmp_risingEdge : BOOL;
END_VAR
(* ENGINEERING_CONTRACT
  Interface contract (per PUB IDs):
  - PUB001: Initial (phase,elapsed,timeout) = (0,0,FALSE) via VAR_INIT.
  - PUB003/PUB004: maxDuration positive INT, finite REALs; no timers/clocks.
  - PUB006/PUB007/PUB008: Per-scan priority: abort > new start rising edge >
    running count. abortBtn TRUE → phase=9 immediately, same-scan start edge
    consumed, re-start requires release+press.
  - PUB009: No abort + new start rising edge → phase=1, elapsed=0, timeout=FALSE;
    start scan not counted.
  - PUB010/PUB011/PUB012: Running state (phase=1 or 2): elapsed increments first,
    then timeout check at updated value (>= maxDuration → phase=3, timeout=TRUE,
    priority over pv/setpoint). Phase transition pv>=setpoint during phase=1
    enters phase=2; phase=2 holds until timeout/abort/new start.
  - PUB013/PUB014: phase=3 (completion) and phase=9 (abort) freeze elapsed and
    timeout until new valid start or abort. No operator acknowledgment.
  Output retention: phase/elapsed/timeout are held in terminal states per S4/N10-S4.
  Same-scan priority: abort evaluated first; start rising edge consumed when abort
    TRUE; timeout check evaluated after elapsed increment and takes priority over
    pv-based phase=2 transition per PUB011.
  Boundary: elapsed>=maxDuration (>= not >) triggers timeout; start scan elapsed=0
    (no increment that scan); trackedPhase preserves same-scan phase context for
    pv evaluation in phase=2 maintenance rule.
*)
BEGIN
    (* Rising edge detection for startBtn (deferred when abort TRUE) *)
    tmp_risingEdge := startBtn AND NOT tmp_startPrev;

    (* Priority 1: abort → phase=9, freeze elapsed & timeout *)
    IF abortBtn THEN
        phase   := 9;
        tmp_phase := phase;
        trackedPhase := phase;
        (* Do NOT update tmp_startPrev; rising edge is consumed per PUB006 *)
    (* Priority 2: new start rising edge → begin new batch *)
    ELSIF tmp_risingEdge THEN
        elapsed     := 0;
        timeout     := FALSE;
        phase       := 1;
        tmp_phase   := phase;
        trackedPhase := phase;
        tmp_startPrev := startBtn;
    (* Priority 3: steady-state running count and phase logic *)
    ELSE
        (* Running state: count one scan, then check timeout, then pv/setpoint *)
        IF (tmp_phase = 1) OR (tmp_phase = 2) THEN
            elapsed := elapsed + 1;
            (* PUB011: timeout check at updated elapsed; priority over pv/setpoint *)
            IF elapsed >= maxDuration THEN
                timeout     := TRUE;
                phase       := 3;
                tmp_phase   := phase;
                trackedPhase := phase;
            ELSIF trackedPhase = 2 OR pv >= setpoint THEN
                phase       := 2;
                tmp_phase   := phase;
                trackedPhase := phase;
            ELSE
                phase       := 1;
                tmp_phase   := phase;
                trackedPhase := phase;
            END_IF;
        ELSE
            (* Idle/completion/abort: hold phase, elapsed, timeout *)
            phase       := tmp_phase;
            trackedPhase := phase;
        END_IF;
        tmp_startPrev := startBtn;
    END_IF;
END_FUNCTION_BLOCK
(* CONTRACT_RULES [] *)

(* ---- self-hard-02.raw_candidate_02.st ---- *)
FUNCTION_BLOCK FB
VAR_INPUT
    startBtn   : BOOL;
    abortBtn   : BOOL;
    setpoint   : REAL;
    pv         : REAL;
    maxDuration: INT;
END_VAR
VAR_OUTPUT
    elapsed : INT := 0;
    phase   : INT := 0;
    timeout : BOOL := FALSE;
END_VAR
VAR
    tmp_startPrev  : BOOL := FALSE;
    tmp_risingEdge : BOOL := FALSE;
    tmp_phase      : INT  := 0;
    trackedPhase   : INT  := 0;
END_VAR
(* ENGINEERING_CONTRACT
  Interface contract (per PUB IDs):
  - PUB001: Initial (phase,elapsed,timeout) = (0,0,FALSE) via VAR_INIT.
  - PUB003/PUB004: maxDuration positive INT, finite REALs; no timers/clocks.
  - PUB006/PUB007/PUB008: Per-scan priority: abort > new start rising edge >
    running count. abortBtn TRUE → phase=9 immediately, same-scan start edge
    consumed, re-start requires release+press.
  - PUB009: No abort + new start rising edge → phase=1, elapsed=0, timeout=FALSE;
    start scan not counted.
  - PUB010/PUB011/PUB012: Running state (phase=1 or 2): elapsed increments first,
    then timeout check at updated value (>= maxDuration → phase=3, timeout=TRUE,
    priority over pv/setpoint). Phase transition pv>=setpoint during phase=1
    enters phase=2; phase=2 holds until timeout/abort/new start.
  - PUB013/PUB014: phase=3 (completion) and phase=9 (abort) freeze elapsed and
    timeout until new valid start or abort. No operator acknowledgment.
  Output retention: phase/elapsed/timeout held in terminal states per S4/N10-S4.
  Same-scan priority: abort evaluated first; start rising edge consumed when abort
    TRUE; timeout check evaluated after elapsed increment and takes priority over
    pv-based phase=2 transition per PUB011.
  Boundary: elapsed>=maxDuration (>=, "reaches") triggers timeout; start scan
    elapsed=0 (no increment that scan); trackedPhase preserves same-scan phase
    context for pv evaluation in phase=2 maintenance rule.
  No unconditional public Boolean latches per CONTRACT_RULES [].
*)
BEGIN
    (* Rising edge detection for startBtn *)
    tmp_risingEdge := startBtn AND NOT tmp_startPrev;

    (* Priority 1: abort → phase=9, freeze elapsed & timeout *)
    IF abortBtn THEN
        phase        := 9;
        tmp_phase    := phase;
        trackedPhase := phase;
    (* Priority 2: new start rising edge → begin new batch *)
    ELSIF tmp_risingEdge THEN
        elapsed      := 0;
        timeout      := FALSE;
        phase        := 1;
        tmp_phase    := phase;
        trackedPhase := phase;
    (* Priority 3: steady-state running count and phase logic *)
    ELSE
        (* Running state: count one scan, then check timeout, then pv/setpoint *)
        IF (tmp_phase = 1) OR (tmp_phase = 2) THEN
            elapsed := elapsed + 1;
            (* PUB011: timeout check at updated elapsed; priority over pv/setpoint *)
            IF elapsed >= maxDuration THEN
                timeout      := TRUE;
                phase        := 3;
                tmp_phase    := phase;
                trackedPhase := phase;
            ELSIF (trackedPhase = 2) OR (pv >= setpoint) THEN
                phase        := 2;
                tmp_phase    := phase;
                trackedPhase := phase;
            ELSE
                phase        := 1;
                tmp_phase    := phase;
                trackedPhase := phase;
            END_IF;
        ELSE
            (* Idle/completion/abort: hold phase, elapsed, timeout *)
            phase        := tmp_phase;
            trackedPhase := phase;
        END_IF;
    END_IF;

    (* Update previous startBtn state for next scan *)
    tmp_startPrev := startBtn;
END_FUNCTION_BLOCK
(* CONTRACT_RULES [] *)

(* ---- self-hard-02.raw_candidate_03.st ---- *)
FUNCTION_BLOCK FB
VAR_INPUT
    startBtn   : BOOL;
    abortBtn   : BOOL;
    setpoint   : REAL;
    pv         : REAL;
    maxDuration: INT;
END_VAR
VAR_OUTPUT
    elapsed : INT := 0;
    phase   : INT := 0;
    timeout : BOOL := FALSE;
END_VAR
VAR
    tmp_startPrev : BOOL := FALSE;
    tmp_phase     : INT  := 0;
END_VAR
VAR
    tmp_risingEdge : BOOL;
END_VAR
(* ENGINEERING_CONTRACT
  Interface contract (per PUB IDs):
  - PUB001: Initial (phase,elapsed,timeout) = (0,0,FALSE) via VAR_INIT.
  - PUB003/PUB004: maxDuration positive INT, finite REALs; no timers/clocks.
  - PUB006/PUB007/PUB008: Per-scan priority: abort > new start rising edge >
    running count. abortBtn TRUE → phase=9 immediately, same-scan start edge
    consumed, re-start requires release+press.
  - PUB009: No abort + new start rising edge → phase=1, elapsed=0, timeout=FALSE;
    start scan not counted.
  - PUB010/PUB011/PUB012: Running state (phase=1 or 2): elapsed increments first,
    then timeout check at updated value (>= maxDuration → phase=3, timeout=TRUE,
    priority over pv/setpoint). Phase transition pv>=setpoint during phase=1
    enters phase=2; phase=2 holds until timeout/abort/new start.
  - PUB013/PUB014: phase=3 (completion) and phase=9 (abort) freeze elapsed and
    timeout until new valid start or abort. No operator acknowledgment.
  Output retention: phase/elapsed/timeout are held in terminal states per S4/N10-S4.
  Same-scan priority: abort evaluated first; start rising edge consumed when abort
    TRUE; timeout check evaluated after elapsed increment and takes priority over
    pv-based phase=2 transition per PUB011.
  Boundary: elapsed>=maxDuration (>= not >) triggers timeout; start scan elapsed=0
    (no increment that scan); tmp_phase preserves same-scan phase context for
    pv evaluation in phase=2 maintenance rule.
*)
BEGIN
    (* Rising edge detection for startBtn (deferred when abort TRUE) *)
    tmp_risingEdge := startBtn AND NOT tmp_startPrev;

    (* Priority 1: abort → phase=9, freeze elapsed & timeout *)
    IF abortBtn THEN
        phase     := 9;
        tmp_phase := phase;
    (* Priority 2: new start rising edge → begin new batch *)
    ELSIF tmp_risingEdge THEN
        elapsed     := 0;
        timeout     := FALSE;
        phase       := 1;
        tmp_phase   := phase;
    (* Priority 3: steady-state running count and phase logic *)
    ELSE
        (* Running state: count one scan, then check timeout, then pv/setpoint *)
        IF (tmp_phase = 1) OR (tmp_phase = 2) THEN
            elapsed := elapsed + 1;
            (* PUB011: timeout check at updated elapsed; priority over pv/setpoint *)
            IF elapsed >= maxDuration THEN
                timeout   := TRUE;
                phase     := 3;
                tmp_phase := phase;
            ELSIF tmp_phase = 2 OR pv >= setpoint THEN
                phase     := 2;
                tmp_phase := phase;
            ELSE
                phase     := 1;
                tmp_phase := phase;
            END_IF;
        ELSE
            (* Idle/completion/abort: hold phase, elapsed, timeout *)
            phase     := tmp_phase;
        END_IF;
        tmp_startPrev := startBtn;
    END_IF;
END_FUNCTION_BLOCK
(* CONTRACT_RULES [] *)

(* ---- self-hard-03.candidate_01.st ---- *)
FUNCTION_BLOCK FB
VAR_INPUT
    pushEn  : BOOL;
    pushItem: INT;
    popEn   : BOOL;
END_VAR
VAR_IN_OUT
    fifo : ARRAY[1..8] OF INT;
END_VAR
VAR_OUTPUT
    count : INT := 0;
    full  : BOOL;
    empty : BOOL;
    head  : INT;
END_VAR
VAR
    pushTrig  : R_TRIG;
    popTrig   : R_TRIG;
    prevCount : INT;
END_VAR

(*
ENGINEERING_CONTRACT
================================================================================
| Output/State  | Activation          | Retention  | Reset      | Priority   |
|---------------|---------------------|------------|------------|------------|
| count         | Rising pushEn OK    | Hold       | Implicit 0 | After pop  |
| full          | count = 8           | Hold       | Implicit   | Same-scan  |
| empty         | count = 0           | Hold       | Implicit   | Same-scan  |
| head          | empty→0 else fifo[1]| Hold       | Implicit   | Same-scan  |
| fifo compact  | After pop+push seq  | Hold       | Implicit   | Pop first  |
--------------------------------------------------------------------------------
PUB001: pushEn rising edge triggers one push per low-to-high transition.
PUB002: popEn rising edge triggers one pop per low-to-high transition.
PUB003: popEn rising edge executes first; removes first item if non-empty.
PUB004: pushEn rising edge executes after pop; appends if count < 8.
PUB005: Full queue with both edges: pop frees slot then push appends.
PUB006: Empty queue with both edges: pop no-op, push adds single item.
PUB007: count = 0..8; full iff count = 8; empty iff count = 0.
PUB008: head = 0 when empty; else head = first item.
PUB009: fifo[1..count] is compact logical queue ordered by pop sequence.
PUB010: fifo[1] = head when non-empty; unspecified beyond count.
--------------------------------------------------------------------------------
CONTRACT_RULES: []
================================================================================
*)
prevCount := count;

pushTrig(CLK := pushEn);
popTrig(CLK := popEn);

IF popTrig.Q AND prevCount > 0 THEN
    FOR 1 TO prevCount - 1 DO
        fifo[i] := fifo[i + 1];
    END_FOR;
    count := prevCount - 1;
ELSE
    count := prevCount;
END_IF;

IF pushTrig.Q THEN
    IF (popTrig.Q AND prevCount > 0) OR (NOT popTrig.Q AND count < 8) THEN
        fifo[count + 1] := pushItem;
        count := count + 1;
    END_IF;
END_IF;

full  := (count = 8);
empty := (count = 0);
head  := SEL(BOOL_TO_INT(empty <> 0), fifo[1], 0);

END_FUNCTION_BLOCK

(* ---- self-hard-03.candidate_02.st ---- *)
FUNCTION_BLOCK FB
VAR_INPUT
    pushEn  : BOOL;
    pushItem: INT;
    popEn   : BOOL;
END_VAR
VAR_IN_OUT
    fifo : ARRAY[1..8] OF INT;
END_VAR
VAR_OUTPUT
    count : INT := 0;
    full  : BOOL;
    empty : BOOL;
    head  : INT;
END_VAR
VAR
    pushTrig  : R_TRIG;
    popTrig   : R_TRIG;
    prevCount : INT;
    tmp_end   : INT;
    tmp_i     : INT;
END_VAR

(*
ENGINEERING_CONTRACT
================================================================================
| Output/State  | Activation          | Retention  | Reset      | Priority   |
|---------------|---------------------|------------|------------|------------|
| count         | Rising pushEn OK    | Hold       | Implicit 0 | After pop  |
| full          | count = 8           | Hold       | Implicit   | Same-scan  |
| empty         | count = 0           | Hold       | Implicit   | Same-scan  |
| head          | empty→0 else fifo[1]| Hold       | Implicit   | Same-scan  |
| fifo compact  | After pop+push seq  | Hold       | Implicit   | Pop first  |
--------------------------------------------------------------------------------
PUB001: pushEn rising edge triggers one push per low-to-high transition.
PUB002: popEn rising edge triggers one pop per low-to-high transition.
PUB003: popEn rising edge executes first; removes first item if non-empty.
PUB004: pushEn rising edge executes after pop; appends if count < 8.
PUB005: Full queue with both edges: pop frees slot then push appends.
PUB006: Empty queue with both edges: pop no-op, push adds single item.
PUB007: count = 0..8; full iff count = 8; empty iff count = 0.
PUB008: head = 0 when empty; else head = first item.
PUB009: fifo[1..count] is compact logical queue ordered by pop sequence.
PUB010: fifo[1] = head when non-empty; unspecified beyond count.
--------------------------------------------------------------------------------
CONTRACT_RULES: []
================================================================================
*)
prevCount := count;

pushTrig(CLK := pushEn);
popTrig(CLK := popEn);

IF popTrig.Q AND prevCount > 0 THEN
    tmp_end := prevCount - 1;
    FOR tmp_i := 1 TO tmp_end DO
        fifo[tmp_i] := fifo[tmp_i + 1];
    END_FOR;
    count := prevCount - 1;
ELSE
    count := prevCount;
END_IF;

IF pushTrig.Q THEN
    IF (popTrig.Q AND prevCount > 0) OR (NOT popTrig.Q AND count < 8) THEN
        fifo[count + 1] := pushItem;
        count := count + 1;
    END_IF;
END_IF;

full  := (count = 8);
empty := (count = 0);
head  := 0;
IF NOT empty THEN
    head := fifo[1];
END_IF;

END_FUNCTION_BLOCK

(* ---- self-hard-03.candidate_03.st ---- *)
FUNCTION_BLOCK FB
VAR_INPUT
    pushEn  : BOOL;
    pushItem: INT;
    popEn   : BOOL;
END_VAR
VAR_IN_OUT
    fifo : ARRAY[1..8] OF INT;
END_VAR
VAR_OUTPUT
    count : INT := 0;
    full  : BOOL;
    empty : BOOL;
    head  : INT;
END_VAR
VAR
    pushTrig  : R_TRIG;
    popTrig   : R_TRIG;
    prevCount : INT;
    tmp_end   : INT;
    tmp_i     : INT;
END_VAR

(*
ENGINEERING_CONTRACT
================================================================================
| Output/State  | Activation          | Retention  | Reset      | Priority   |
|---------------|---------------------|------------|------------|------------|
| count         | pushEn=1 AND cond   | Hold       | Implicit 0 | After pop  |
| full          | count = 8           | Hold       | Implicit   | Same-scan  |
| empty         | count = 0           | Hold       | Implicit   | Same-scan  |
| head          | empty→0 else fifo[1]| Hold       | Implicit   | Same-scan  |
| fifo compact  | After pop+push seq  | Hold       | Implicit   | Pop first  |
--------------------------------------------------------------------------------
PUB001: pushEn rising edge triggers one push per low-to-high transition.
PUB002: popEn rising edge triggers one pop per low-to-high transition.
PUB003: popEn rising edge executes first; removes first item if non-empty.
PUB004: pushEn rising edge executes after pop; appends if count < 8.
PUB005: Full queue with both edges: pop frees slot then push appends.
PUB006: Empty queue with both edges: pop no-op, push adds single item.
PUB007: count = 0..8; full iff count = 8; empty iff count = 0.
PUB008: head = 0 when empty; else head = first item.
PUB009: fifo[1..count] is compact logical queue ordered by pop sequence.
PUB010: fifo[1] = head when non-empty; unspecified beyond count.
--------------------------------------------------------------------------------
CONTRACT_RULES: []
================================================================================
*)
prevCount := count;

pushTrig(CLK := pushEn);
popTrig(CLK := popEn);

IF popTrig.Q AND prevCount > 0 THEN
    tmp_end := prevCount - 1;
    FOR tmp_i := 1 TO tmp_end DO
        fifo[tmp_i] := fifo[tmp_i + 1];
    END_FOR;
    count := prevCount - 1;
ELSE
    count := prevCount;
END_IF;

IF pushEn AND ((popTrig.Q AND prevCount > 0) OR (NOT (prevCount = 0 AND popTrig.Q) AND count < 8)) THEN
    fifo[count + 1] := pushItem;
    count := count + 1;
END_IF;

full  := (count = 8);
empty := (count = 0);
head  := 0;
IF NOT empty THEN
    head := fifo[1];
END_IF;

END_FUNCTION_BLOCK

(* ---- self-hard-03.candidate_04.st ---- *)
FUNCTION_BLOCK FB
VAR_INPUT
    pushEn  : BOOL;
    pushItem: INT;
    popEn   : BOOL;
END_VAR
VAR_IN_OUT
    fifo : ARRAY[1..8] OF INT;
END_VAR
VAR_OUTPUT
    count : INT := 0;
    full  : BOOL;
    empty : BOOL;
    head  : INT;
END_VAR
VAR
    pushTrig  : R_TRIG;
    popTrig   : R_TRIG;
    prevCount : INT;
    tmp_end   : INT;
    tmp_i     : INT;
END_VAR

(*
ENGINEERING_CONTRACT
================================================================================
| Output/State  | Activation          | Retention  | Reset      | Priority   |
|---------------|---------------------|------------|------------|------------|
| count         | Rising pushEn OK    | Hold       | Implicit 0 | After pop  |
| full          | count = 8           | Hold       | Implicit   | Same-scan  |
| empty         | count = 0           | Hold       | Implicit   | Same-scan  |
| head          | empty→0 else fifo[1]| Hold       | Implicit   | Same-scan  |
| fifo compact  | After pop+push seq  | Hold       | Implicit   | Pop first  |
--------------------------------------------------------------------------------
PUB001: pushEn rising edge triggers one push per low-to-high transition.
PUB002: popEn rising edge triggers one pop per low-to-high transition.
PUB003: popEn rising edge executes first; removes first item if non-empty.
PUB004: pushEn rising edge executes after pop; appends if count < 8.
PUB005: Full queue with both edges: pop frees slot then push appends.
PUB006: Empty queue with both edges: pop no-op, push adds single item.
PUB007: count = 0..8; full iff count = 8; empty iff count = 0.
PUB008: head = 0 when empty; else head = first item.
PUB009: fifo[1..count] is compact logical queue ordered by pop sequence.
PUB010: fifo[1] = head when non-empty; unspecified beyond count.
--------------------------------------------------------------------------------
CONTRACT_RULES: []
================================================================================
*)
prevCount := count;

pushTrig(CLK := pushEn);
popTrig(CLK := popEn);

IF popTrig.Q AND prevCount > 0 THEN
    tmp_end := prevCount - 1;
    FOR tmp_i := 1 TO tmp_end DO
        fifo[tmp_i] := fifo[tmp_i + 1];
    END_FOR;
    count := prevCount - 1;
ELSE
    count := prevCount;
END_IF;

IF pushTrig.Q THEN
    IF popTrig.Q OR (count < 8) THEN
        fifo[count + 1] := pushItem;
        count := count + 1;
    END_IF;
END_IF;

full  := (count = 8);
empty := (count = 0);
head  := 0;
IF NOT empty THEN
    head := fifo[1];
END_IF;

END_FUNCTION_BLOCK

(* ---- self-hard-03.raw_candidate_01.st ---- *)
FUNCTION_BLOCK FB
VAR_INPUT
    pushEn  : BOOL;
    pushItem: INT;
    popEn   : BOOL;
END_VAR
VAR_IN_OUT
    fifo : ARRAY[1..8] OF INT;
END_VAR
VAR_OUTPUT
    count : INT := 0;
    full  : BOOL;
    empty : BOOL;
    head  : INT;
END_VAR
VAR
    pushTrig  : R_TRIG;
    popTrig   : R_TRIG;
    prevCount : INT;
END_VAR

(*
ENGINEERING_CONTRACT
================================================================================
| Output/State  | Activation          | Retention  | Reset      | Priority   |
|---------------|---------------------|------------|------------|------------|
| count         | Rising pushEn OK    | Hold       | Implicit 0 | After pop  |
| full          | count = 8           | Hold       | Implicit   | Same-scan  |
| empty         | count = 0           | Hold       | Implicit   | Same-scan  |
| head          | empty→0 else fifo[1]| Hold       | Implicit   | Same-scan  |
| fifo compact  | After pop+push seq  | Hold       | Implicit   | Pop first  |
--------------------------------------------------------------------------------
PUB001: pushEn rising edge triggers one push per low-to-high transition.
PUB002: popEn rising edge triggers one pop per low-to-high transition.
PUB003: popEn rising edge executes first; removes first item if non-empty.
PUB004: pushEn rising edge executes after pop; appends if count < 8.
PUB005: Full queue with both edges: pop frees slot then push appends.
PUB006: Empty queue with both edges: pop no-op, push adds single item.
PUB007: count = 0..8; full iff count = 8; empty iff count = 0.
PUB008: head = 0 when empty; else head = first item.
PUB009: fifo[1..count] is compact logical queue ordered by pop sequence.
PUB010: fifo[1] = head when non-empty; unspecified beyond count.
--------------------------------------------------------------------------------
CONTRACT_RULES: []
================================================================================
*)
prevCount := count;

pushTrig(CLK := pushEn);
popTrig(CLK := popEn);

IF popTrig.Q AND prevCount > 0 THEN
    FOR 1 TO prevCount - 1 DO
        fifo[i] := fifo[i + 1];
    END_FOR;
    count := prevCount - 1;
ELSE
    count := prevCount;
END_IF;

IF pushTrig.Q THEN
    IF (popTrig.Q AND prevCount > 0) OR (NOT popTrig.Q AND count < 8) THEN
        fifo[count + 1] := pushItem;
        count := count + 1;
    END_IF;
END_IF;

full  := (count = 8);
empty := (count = 0);
head  := SEL(BOOL_TO_INT(empty <> 0), fifo[1], 0);

END_FUNCTION_BLOCK

(* ---- self-hard-03.raw_candidate_02.st ---- *)
FUNCTION_BLOCK FB
VAR_INPUT
    pushEn  : BOOL;
    pushItem: INT;
    popEn   : BOOL;
END_VAR
VAR_IN_OUT
    fifo : ARRAY[1..8] OF INT;
END_VAR
VAR_OUTPUT
    count : INT := 0;
    full  : BOOL;
    empty : BOOL;
    head  : INT;
END_VAR
VAR
    pushTrig  : R_TRIG;
    popTrig   : R_TRIG;
    prevCount : INT;
    tmp_end   : INT;
    tmp_i     : INT;
END_VAR

(*
ENGINEERING_CONTRACT
================================================================================
| Output/State  | Activation          | Retention  | Reset      | Priority   |
|---------------|---------------------|------------|------------|------------|
| count         | Rising pushEn OK    | Hold       | Implicit 0 | After pop  |
| full          | count = 8           | Hold       | Implicit   | Same-scan  |
| empty         | count = 0           | Hold       | Implicit   | Same-scan  |
| head          | empty→0 else fifo[1]| Hold       | Implicit   | Same-scan  |
| fifo compact  | After pop+push seq  | Hold       | Implicit   | Pop first  |
--------------------------------------------------------------------------------
PUB001: pushEn rising edge triggers one push per low-to-high transition.
PUB002: popEn rising edge triggers one pop per low-to-high transition.
PUB003: popEn rising edge executes first; removes first item if non-empty.
PUB004: pushEn rising edge executes after pop; appends if count < 8.
PUB005: Full queue with both edges: pop frees slot then push appends.
PUB006: Empty queue with both edges: pop no-op, push adds single item.
PUB007: count = 0..8; full iff count = 8; empty iff count = 0.
PUB008: head = 0 when empty; else head = first item.
PUB009: fifo[1..count] is compact logical queue ordered by pop sequence.
PUB010: fifo[1] = head when non-empty; unspecified beyond count.
--------------------------------------------------------------------------------
CONTRACT_RULES: []
================================================================================
*)
prevCount := count;

pushTrig(CLK := pushEn);
popTrig(CLK := popEn);

IF popTrig.Q AND prevCount > 0 THEN
    tmp_end := prevCount - 1;
    FOR tmp_i := 1 TO tmp_end DO
        fifo[tmp_i] := fifo[tmp_i + 1];
    END_FOR;
    count := prevCount - 1;
ELSE
    count := prevCount;
END_IF;

IF pushTrig.Q THEN
    IF (popTrig.Q AND prevCount > 0) OR (NOT popTrig.Q AND count < 8) THEN
        fifo[count + 1] := pushItem;
        count := count + 1;
    END_IF;
END_IF;

full  := (count = 8);
empty := (count = 0);
head  := 0;
IF NOT empty THEN
    head := fifo[1];
END_IF;

END_FUNCTION_BLOCK

(* ---- self-hard-03.raw_candidate_03.st ---- *)
FUNCTION_BLOCK FB
VAR_INPUT
    pushEn  : BOOL;
    pushItem: INT;
    popEn   : BOOL;
END_VAR
VAR_IN_OUT
    fifo : ARRAY[1..8] OF INT;
END_VAR
VAR_OUTPUT
    count : INT := 0;
    full  : BOOL;
    empty : BOOL;
    head  : INT;
END_VAR
VAR
    pushTrig  : R_TRIG;
    popTrig   : R_TRIG;
    prevCount : INT;
    tmp_end   : INT;
    tmp_i     : INT;
END_VAR

(*
ENGINEERING_CONTRACT
================================================================================
| Output/State  | Activation          | Retention  | Reset      | Priority   |
|---------------|---------------------|------------|------------|------------|
| count         | pushEn=1 AND cond   | Hold       | Implicit 0 | After pop  |
| full          | count = 8           | Hold       | Implicit   | Same-scan  |
| empty         | count = 0           | Hold       | Implicit   | Same-scan  |
| head          | empty→0 else fifo[1]| Hold       | Implicit   | Same-scan  |
| fifo compact  | After pop+push seq  | Hold       | Implicit   | Pop first  |
--------------------------------------------------------------------------------
PUB001: pushEn rising edge triggers one push per low-to-high transition.
PUB002: popEn rising edge triggers one pop per low-to-high transition.
PUB003: popEn rising edge executes first; removes first item if non-empty.
PUB004: pushEn rising edge executes after pop; appends if count < 8.
PUB005: Full queue with both edges: pop frees slot then push appends.
PUB006: Empty queue with both edges: pop no-op, push adds single item.
PUB007: count = 0..8; full iff count = 8; empty iff count = 0.
PUB008: head = 0 when empty; else head = first item.
PUB009: fifo[1..count] is compact logical queue ordered by pop sequence.
PUB010: fifo[1] = head when non-empty; unspecified beyond count.
--------------------------------------------------------------------------------
CONTRACT_RULES: []
================================================================================
*)
prevCount := count;

pushTrig(CLK := pushEn);
popTrig(CLK := popEn);

IF popTrig.Q AND prevCount > 0 THEN
    tmp_end := prevCount - 1;
    FOR tmp_i := 1 TO tmp_end DO
        fifo[tmp_i] := fifo[tmp_i + 1];
    END_FOR;
    count := prevCount - 1;
ELSE
    count := prevCount;
END_IF;

IF pushEn AND ((popTrig.Q AND prevCount > 0) OR (NOT (prevCount = 0 AND popTrig.Q) AND count < 8)) THEN
    fifo[count + 1] := pushItem;
    count := count + 1;
END_IF;

full  := (count = 8);
empty := (count = 0);
head  := 0;
IF NOT empty THEN
    head := fifo[1];
END_IF;

END_FUNCTION_BLOCK

(* ---- self-hard-03.raw_candidate_04.st ---- *)
FUNCTION_BLOCK FB
VAR_INPUT
    pushEn  : BOOL;
    pushItem: INT;
    popEn   : BOOL;
END_VAR
VAR_IN_OUT
    fifo : ARRAY[1..8] OF INT;
END_VAR
VAR_OUTPUT
    count : INT := 0;
    full  : BOOL;
    empty : BOOL;
    head  : INT;
END_VAR
VAR
    pushTrig  : R_TRIG;
    popTrig   : R_TRIG;
    prevCount : INT;
    tmp_end   : INT;
    tmp_i     : INT;
END_VAR

(*
ENGINEERING_CONTRACT
================================================================================
| Output/State  | Activation          | Retention  | Reset      | Priority   |
|---------------|---------------------|------------|------------|------------|
| count         | Rising pushEn OK    | Hold       | Implicit 0 | After pop  |
| full          | count = 8           | Hold       | Implicit   | Same-scan  |
| empty         | count = 0           | Hold       | Implicit   | Same-scan  |
| head          | empty→0 else fifo[1]| Hold       | Implicit   | Same-scan  |
| fifo compact  | After pop+push seq  | Hold       | Implicit   | Pop first  |
--------------------------------------------------------------------------------
PUB001: pushEn rising edge triggers one push per low-to-high transition.
PUB002: popEn rising edge triggers one pop per low-to-high transition.
PUB003: popEn rising edge executes first; removes first item if non-empty.
PUB004: pushEn rising edge executes after pop; appends if count < 8.
PUB005: Full queue with both edges: pop frees slot then push appends.
PUB006: Empty queue with both edges: pop no-op, push adds single item.
PUB007: count = 0..8; full iff count = 8; empty iff count = 0.
PUB008: head = 0 when empty; else head = first item.
PUB009: fifo[1..count] is compact logical queue ordered by pop sequence.
PUB010: fifo[1] = head when non-empty; unspecified beyond count.
--------------------------------------------------------------------------------
CONTRACT_RULES: []
================================================================================
*)
prevCount := count;

pushTrig(CLK := pushEn);
popTrig(CLK := popEn);

IF popTrig.Q AND prevCount > 0 THEN
    tmp_end := prevCount - 1;
    FOR tmp_i := 1 TO tmp_end DO
        fifo[tmp_i] := fifo[tmp_i + 1];
    END_FOR;
    count := prevCount - 1;
ELSE
    count := prevCount;
END_IF;

IF pushTrig.Q THEN
    IF popTrig.Q OR (count < 8) THEN
        fifo[count + 1] := pushItem;
        count := count + 1;
    END_IF;
END_IF;

full  := (count = 8);
empty := (count = 0);
head  := 0;
IF NOT empty THEN
    head := fifo[1];
END_IF;

END_FUNCTION_BLOCK

(* ---- self-hard-04.candidate_01.st ---- *)
FUNCTION_BLOCK FB
VAR_OUTPUT
    leadPump : INT := 0;
    lagPump : INT := 0;
    runningCount : INT := 0;
END_VAR
VAR_INPUT
    demand : INT;
    runHours : ARRAY[1..5] OF LINT;
    rotated : BOOL;
END_VAR
VAR
    tmp_prevLead : INT := 0;
    tmp_prevRunning : INT := 0;
    tmp_selectLag : BOOL := FALSE;
    tmp_newLead : INT;
    minHours : LINT;
    i : INT;
END_VAR
VAR_TEMP
    newLag : INT;
END_VAR
(*
ENGINEERING_CONTRACT:
  [S1] runningCount = CLAMP(demand, 0, 5). PUB001/PUB011
  [S2] demand=0→leadPump=lagPump=0; demand=1→lagPump=0; demand≥2→leadPump≠lagPump, both 1..5. PUB002/PUB012
  [S3] Lead-change requires old lead hours > new lead hours + 50. PUB036
  [S4] Hysteresis: rotated=TRUE AND runHours[lead] > minHours + 50 → rotate to min-hours pump. PUB026/PUB027
  [S5] Lag pump selected ONLY on: initial, lead change, runningCount increase. PUB005/PUB031
  [S6] Initial lead selection: min (runHours, pump#). PUB028
  [S7] Lag pump: min (runHours, pump#) excluding lead pump. PUB029
  [S8] Demand=0 clears lead/lag immediately; next positive demand triggers fresh selection. PUB033/PUB034
  [S9] First FB invocation initializes all outputs to 0 (VAR_INIT). PUB041
  No edge detection on rotated; it is level-triggered. PUB026
  Array bounds: 1..5 only. PUB042
*)
(* CONTRACT_RULES [] *)

tmp_prevLead := leadPump;
tmp_prevRunning := runningCount;
tmp_selectLag := FALSE;

IF demand <= 0 THEN
    runningCount := 0;
    leadPump := 0;
    lagPump := 0;
ELSIF leadPump = 0 THEN
    runningCount := demand;
    tmp_newLead := 1;
    FOR i := 2 TO 5 DO
        IF runHours[i] < runHours[tmp_newLead] OR (runHours[i] = runHours[tmp_newLead] AND i < tmp_newLead) THEN
            tmp_newLead := i;
        END_IF;
    END_FOR;
    leadPump := tmp_newLead;
    tmp_selectLag := TRUE;
    IF demand >= 2 THEN
        newLag := 0;
        FOR i := 1 TO 5 DO
            IF i <> leadPump THEN
                IF newLag = 0 OR runHours[i] < runHours[newLag] OR (runHours[i] = runHours[newLag] AND i < newLag) THEN
                    newLag := i;
                END_IF;
            END_IF;
        END_FOR;
        lagPump := newLag;
    ELSE
        lagPump := 0;
    END_IF;
ELSE
    runningCount := demand;
    IF rotated AND runHours[leadPump] > minHours + 50 THEN
        tmp_newLead := 1;
        FOR i := 2 TO 5 DO
            IF runHours[i] < runHours[tmp_newLead] OR (runHours[i] = runHours[tmp_newLead] AND i < tmp_newLead) THEN
                tmp_newLead := i;
            END_IF;
        END_FOR;
        leadPump := tmp_newLead;
        tmp_selectLag := TRUE;
    END_IF;
    IF demand > tmp_prevRunning THEN
        tmp_newLead := 1;
        FOR i := 2 TO 5 DO
            IF runHours[i] < runHours[tmp_newLead] OR (runHours[i] = runHours[tmp_newLead] AND i < tmp_newLead) THEN
                tmp_newLead := i;
            END_IF;
        END_FOR;
        leadPump := tmp_newLead;
        tmp_selectLag := TRUE;
    END_IF;
    IF tmp_selectLag THEN
        IF demand >= 2 THEN
            newLag := 0;
            FOR i := 1 TO 5 DO
                IF i <> leadPump THEN
                    IF newLag = 0 OR runHours[i] < runHours[newLag] OR (runHours[i] = runHours[newLag] AND i < newLag) THEN
                        newLag := i;
                    END_IF;
                END_IF;
            END_FOR;
            lagPump := newLag;
        ELSE
            lagPump := 0;
        END_IF;
    END_IF;
END_IF;

minHours := runHours[1];
FOR i := 2 TO 5 DO
    IF runHours[i] < minHours THEN
        minHours := runHours[i];
    END_IF;
END_FOR;
END_FUNCTION_BLOCK

(* ---- self-hard-04.candidate_02.st ---- *)
FUNCTION_BLOCK FB
VAR_OUTPUT
    leadPump : INT := 0;
    lagPump : INT := 0;
    runningCount : INT := 0;
END_VAR
VAR_INPUT
    demand : INT;
    runHours : ARRAY[1..5] OF LINT;
    rotated : BOOL;
END_VAR
VAR
    tmp_prevLead : INT := 0;
    tmp_prevRunning : INT := 0;
    tmp_selectLag : BOOL := FALSE;
    tmp_newLead : INT;
    tmp_minOther : LINT;
    i : INT;
END_VAR
VAR_TEMP
    newLag : INT;
    clippedDemand : INT;
END_VAR
(*
ENGINEERING_CONTRACT:
  [S1] runningCount = CLAMP(demand, 0, 5). PUB001/PUB011
  [S2] demand=0→leadPump=lagPump=0; demand=1→lagPump=0; demand≥2→leadPump≠lagPump, both 1..5. PUB002/PUB012
  [S3] Lead-change requires old lead hours > new lead hours + 50. PUB036
  [S4] Hysteresis: rotated=TRUE AND runHours[lead] > minOther + 50 → rotate to min-other pump. PUB026/PUB027
  [S5] Lag pump selected ONLY on: initial, lead change, runningCount increase. PUB005/PUB031
  [S6] Initial lead selection: min (runHours, pump#). PUB028
  [S7] Lag pump: min (runHours, pump#) excluding lead pump. PUB029
  [S8] Demand=0 clears lead/lag immediately; next positive demand triggers fresh selection. PUB033/PUB034
  [S9] First FB invocation initializes all outputs to 0 (VAR_INIT). PUB041
  No edge detection on rotated; it is level-triggered. PUB026
  Array bounds: 1..5 only. PUB042
*)
(* CONTRACT_RULES [] *)

clippedDemand := demand;
IF clippedDemand < 0 THEN
    clippedDemand := 0;
ELSIF clippedDemand > 5 THEN
    clippedDemand := 5;
END_IF;

tmp_prevLead := leadPump;
tmp_prevRunning := runningCount;
tmp_selectLag := FALSE;

IF clippedDemand = 0 THEN
    runningCount := 0;
    leadPump := 0;
    lagPump := 0;
ELSIF leadPump = 0 THEN
    runningCount := clippedDemand;
    tmp_newLead := 1;
    FOR i := 2 TO 5 DO
        IF runHours[i] < runHours[tmp_newLead] OR (runHours[i] = runHours[tmp_newLead] AND i < tmp_newLead) THEN
            tmp_newLead := i;
        END_IF;
    END_FOR;
    leadPump := tmp_newLead;
    tmp_selectLag := TRUE;
    IF clippedDemand >= 2 THEN
        newLag := 0;
        FOR i := 1 TO 5 DO
            IF i <> leadPump THEN
                IF newLag = 0 OR runHours[i] < runHours[newLag] OR (runHours[i] = runHours[newLag] AND i < newLag) THEN
                    newLag := i;
                END_IF;
            END_IF;
        END_FOR;
        lagPump := newLag;
    ELSE
        lagPump := 0;
    END_IF;
ELSE
    runningCount := clippedDemand;
    tmp_minOther := 9223372036854775807; // LINT_MAX approximation
    FOR i := 1 TO 5 DO
        IF i <> leadPump AND runHours[i] < tmp_minOther THEN
            tmp_minOther := runHours[i];
        END_IF;
    END_FOR;
    IF rotated AND runHours[leadPump] > tmp_minOther + 50 THEN
        tmp_newLead := 1;
        FOR i := 2 TO 5 DO
            IF runHours[i] < runHours[tmp_newLead] OR (runHours[i] = runHours[tmp_newLead] AND i < tmp_newLead) THEN
                tmp_newLead := i;
            END_IF;
        END_FOR;
        leadPump := tmp_newLead;
        tmp_selectLag := TRUE;
    END_IF;
    IF clippedDemand > tmp_prevRunning THEN
        tmp_newLead := 1;
        FOR i := 2 TO 5 DO
            IF runHours[i] < runHours[tmp_newLead] OR (runHours[i] = runHours[tmp_newLead] AND i < tmp_newLead) THEN
                tmp_newLead := i;
            END_IF;
        END_FOR;
        leadPump := tmp_newLead;
        tmp_selectLag := TRUE;
    END_IF;
    IF tmp_selectLag THEN
        IF clippedDemand >= 2 THEN
            newLag := 0;
            FOR i := 1 TO 5 DO
                IF i <> leadPump THEN
                    IF newLag = 0 OR runHours[i] < runHours[newLag] OR (runHours[i] = runHours[newLag] AND i < newLag) THEN
                        newLag := i;
                    END_IF;
                END_IF;
            END_FOR;
            lagPump := newLag;
        ELSE
            lagPump := 0;
        END_IF;
    END_IF;
END_IF;
END_FUNCTION_BLOCK

(* ---- self-hard-04.candidate_03.st ---- *)
FUNCTION_BLOCK FB
VAR_OUTPUT
    leadPump : INT := 0;
    lagPump : INT := 0;
    runningCount : INT := 0;
END_VAR
VAR_INPUT
    demand : INT;
    runHours : ARRAY[1..5] OF LINT;
    rotated : BOOL;
END_VAR
VAR
    tmp_prevLead : INT := 0;
    tmp_prevRunning : INT := 0;
    tmp_selectLag : BOOL := FALSE;
    tmp_newLead : INT;
    minHours : LINT;
    i : INT;
    tmp_demand : INT;
END_VAR
VAR_TEMP
    newLag : INT;
END_VAR
(*
ENGINEERING_CONTRACT:
  [S1] runningCount = CLAMP(demand, 0, 5). PUB001/PUB011
  [S2] demand=0→leadPump=lagPump=0; demand=1→lagPump=0; demand≥2→leadPump≠lagPump, both 1..5. PUB002/PUB012
  [S3] Lead-change requires old lead hours > new lead hours + 50. PUB036
  [S4] Hysteresis: rotated=TRUE AND runHours[lead] > minHours + 50 → rotate to min-hours pump. PUB026/PUB027
  [S5] Lag pump selected ONLY on: initial, lead change, runningCount increase. PUB005/PUB031
  [S6] Initial lead selection: min (runHours, pump#). PUB028
  [S7] Lag pump: min (runHours, pump#) excluding lead pump. PUB029
  [S8] Demand=0 clears lead/lag immediately; next positive demand triggers fresh selection. PUB033/PUB034
  [S9] First FB invocation initializes all outputs to 0 (VAR_INIT). PUB041
  No edge detection on rotated; it is level-triggered. PUB026
  Array bounds: 1..5 only. PUB042
*)
(* CONTRACT_RULES [] *)

tmp_prevLead := leadPump;
tmp_prevRunning := runningCount;
tmp_selectLag := FALSE;

IF demand < 0 THEN
    tmp_demand := 0;
ELSIF demand > 5 THEN
    tmp_demand := 5;
ELSE
    tmp_demand := demand;
END_IF;

minHours := runHours[1];
FOR i := 2 TO 5 DO
    IF runHours[i] < minHours THEN
        minHours := runHours[i];
    END_IF;
END_FOR;

IF tmp_demand <= 0 THEN
    runningCount := 0;
    leadPump := 0;
    lagPump := 0;
ELSIF tmp_prevLead = 0 THEN
    runningCount := tmp_demand;
    tmp_newLead := 1;
    FOR i := 2 TO 5 DO
        IF runHours[i] < runHours[tmp_newLead] OR (runHours[i] = runHours[tmp_newLead] AND i < tmp_newLead) THEN
            tmp_newLead := i;
        END_IF;
    END_FOR;
    leadPump := tmp_newLead;
    tmp_selectLag := TRUE;
    IF tmp_demand >= 2 THEN
        newLag := 0;
        FOR i := 1 TO 5 DO
            IF i <> leadPump THEN
                IF newLag = 0 OR runHours[i] < runHours[newLag] OR (runHours[i] = runHours[newLag] AND i < newLag) THEN
                    newLag := i;
                END_IF;
            END_IF;
        END_FOR;
        lagPump := newLag;
    ELSE
        lagPump := 0;
    END_IF;
ELSE
    runningCount := tmp_demand;
    IF rotated AND runHours[leadPump] > minHours + 50 THEN
        tmp_newLead := 1;
        FOR i := 2 TO 5 DO
            IF runHours[i] < runHours[tmp_newLead] OR (runHours[i] = runHours[tmp_newLead] AND i < tmp_newLead) THEN
                tmp_newLead := i;
            END_IF;
        END_FOR;
        leadPump := tmp_newLead;
        tmp_selectLag := TRUE;
    END_IF;
    IF tmp_demand > tmp_prevRunning THEN
        tmp_newLead := 1;
        FOR i := 2 TO 5 DO
            IF runHours[i] < runHours[tmp_newLead] OR (runHours[i] = runHours[tmp_newLead] AND i < tmp_newLead) THEN
                tmp_newLead := i;
            END_IF;
        END_FOR;
        leadPump := tmp_newLead;
        tmp_selectLag := TRUE;
    END_IF;
    IF tmp_selectLag THEN
        IF tmp_demand >= 2 THEN
            newLag := 0;
            FOR i := 1 TO 5 DO
                IF i <> leadPump THEN
                    IF newLag = 0 OR runHours[i] < runHours[newLag] OR (runHours[i] = runHours[newLag] AND i < newLag) THEN
                        newLag := i;
                    END_IF;
                END_IF;
            END_FOR;
            lagPump := newLag;
        ELSE
            lagPump := 0;
        END_IF;
    END_IF;
END_IF;
END_FUNCTION_BLOCK

(* ---- self-hard-04.candidate_04.st ---- *)
FUNCTION_BLOCK FB
VAR_OUTPUT
    leadPump : INT := 0;
    lagPump : INT := 0;
    runningCount : INT := 0;
END_VAR
VAR_INPUT
    demand : INT;
    runHours : ARRAY[1..5] OF LINT;
    rotated : BOOL;
END_VAR
VAR
    tmp_prevLead : INT := 0;
    tmp_prevRunning : INT := 0;
    tmp_selectLag : BOOL := FALSE;
    tmp_newLead : INT;
    minHours : LINT;
    i : INT;
END_VAR
VAR_TEMP
    newLag : INT;
END_VAR
(*
ENGINEERING_CONTRACT:
  [S1] runningCount = CLAMP(demand, 0, 5). PUB001/PUB011
  [S2] demand=0→leadPump=lagPump=0; demand=1→lagPump=0; demand≥2→leadPump≠lagPump, both 1..5. PUB002/PUB012
  [S3] Lead-change requires old lead hours > new lead hours + 50. PUB036
  [S4] Hysteresis: rotated=TRUE AND runHours[lead] > minHours + 50 → rotate to min-hours pump. PUB026/PUB027
  [S5] Lag pump selected ONLY on: initial, lead change, runningCount increase. PUB005/PUB031
  [S6] Initial lead selection: min (runHours, pump#). PUB028
  [S7] Lag pump: min (runHours, pump#) excluding lead pump. PUB029
  [S8] Demand=0 clears lead/lag immediately; next positive demand triggers fresh selection. PUB033/PUB034
  [S9] First FB invocation initializes all outputs to 0 (VAR_INIT). PUB041
  No edge detection on rotated; it is level-triggered. PUB026
  Array bounds: 1..5 only. PUB042
*)
(* CONTRACT_RULES [] *)

tmp_prevLead := leadPump;
tmp_prevRunning := runningCount;
tmp_selectLag := FALSE;

minHours := runHours[1];
FOR i := 2 TO 5 DO
    IF runHours[i] < minHours THEN
        minHours := runHours[i];
    END_IF;
END_FOR;

IF demand <= 0 THEN
    runningCount := 0;
    leadPump := 0;
    lagPump := 0;
ELSIF leadPump = 0 THEN
    runningCount := demand;
    IF demand > 5 THEN
        runningCount := 5;
    ELSIF demand < 0 THEN
        runningCount := 0;
    END_IF;
    tmp_newLead := 1;
    FOR i := 2 TO 5 DO
        IF runHours[i] < runHours[tmp_newLead] OR (runHours[i] = runHours[tmp_newLead] AND i < tmp_newLead) THEN
            tmp_newLead := i;
        END_IF;
    END_FOR;
    leadPump := tmp_newLead;
    tmp_selectLag := TRUE;
    IF demand >= 2 THEN
        newLag := 0;
        FOR i := 1 TO 5 DO
            IF i <> leadPump THEN
                IF newLag = 0 OR runHours[i] < runHours[newLag] OR (runHours[i] = runHours[newLag] AND i < newLag) THEN
                    newLag := i;
                END_IF;
            END_IF;
        END_FOR;
        lagPump := newLag;
    ELSE
        lagPump := 0;
    END_IF;
ELSE
    IF demand > 5 THEN
        runningCount := 5;
    ELSIF demand < 0 THEN
        runningCount := 0;
    ELSE
        runningCount := demand;
    END_IF;
    IF rotated AND runHours[leadPump] > minHours + 50 THEN
        tmp_newLead := 1;
        FOR i := 2 TO 5 DO
            IF runHours[i] < runHours[tmp_newLead] OR (runHours[i] = runHours[tmp_newLead] AND i < tmp_newLead) THEN
                tmp_newLead := i;
            END_IF;
        END_FOR;
        leadPump := tmp_newLead;
        tmp_selectLag := TRUE;
    END_IF;
    IF demand > tmp_prevRunning THEN
        tmp_newLead := 1;
        FOR i := 2 TO 5 DO
            IF runHours[i] < runHours[tmp_newLead] OR (runHours[i] = runHours[tmp_newLead] AND i < tmp_newLead) THEN
                tmp_newLead := i;
            END_IF;
        END_FOR;
        leadPump := tmp_newLead;
        tmp_selectLag := TRUE;
    END_IF;
    IF tmp_selectLag THEN
        IF demand >= 2 THEN
            newLag := 0;
            FOR i := 1 TO 5 DO
                IF i <> leadPump THEN
                    IF newLag = 0 OR runHours[i] < runHours[newLag] OR (runHours[i] = runHours[newLag] AND i < newLag) THEN
                        newLag := i;
                    END_IF;
                END_IF;
            END_FOR;
            lagPump := newLag;
        ELSE
            lagPump := 0;
        END_IF;
    END_IF;
END_IF;
END_FUNCTION_BLOCK

(* ---- self-hard-04.raw_candidate_01.st ---- *)
FUNCTION_BLOCK FB
VAR_OUTPUT
    leadPump : INT := 0;
    lagPump : INT := 0;
    runningCount : INT := 0;
END_VAR
VAR_INPUT
    demand : INT;
    runHours : ARRAY[1..5] OF LINT;
    rotated : BOOL;
END_VAR
VAR
    tmp_prevLead : INT := 0;
    tmp_prevRunning : INT := 0;
    tmp_selectLag : BOOL := FALSE;
    tmp_newLead : INT;
    minHours : LINT;
    i : INT;
END_VAR
VAR_TEMP
    newLag : INT;
END_VAR
(*
ENGINEERING_CONTRACT:
  [S1] runningCount = CLAMP(demand, 0, 5). PUB001/PUB011
  [S2] demand=0→leadPump=lagPump=0; demand=1→lagPump=0; demand≥2→leadPump≠lagPump, both 1..5. PUB002/PUB012
  [S3] Lead-change requires old lead hours > new lead hours + 50. PUB036
  [S4] Hysteresis: rotated=TRUE AND runHours[lead] > minHours + 50 → rotate to min-hours pump. PUB026/PUB027
  [S5] Lag pump selected ONLY on: initial, lead change, runningCount increase. PUB005/PUB031
  [S6] Initial lead selection: min (runHours, pump#). PUB028
  [S7] Lag pump: min (runHours, pump#) excluding lead pump. PUB029
  [S8] Demand=0 clears lead/lag immediately; next positive demand triggers fresh selection. PUB033/PUB034
  [S9] First FB invocation initializes all outputs to 0 (VAR_INIT). PUB041
  No edge detection on rotated; it is level-triggered. PUB026
  Array bounds: 1..5 only. PUB042
*)
(* CONTRACT_RULES [] *)

tmp_prevLead := leadPump;
tmp_prevRunning := runningCount;
tmp_selectLag := FALSE;

IF demand <= 0 THEN
    runningCount := 0;
    leadPump := 0;
    lagPump := 0;
ELSIF leadPump = 0 THEN
    runningCount := demand;
    tmp_newLead := 1;
    FOR i := 2 TO 5 DO
        IF runHours[i] < runHours[tmp_newLead] OR (runHours[i] = runHours[tmp_newLead] AND i < tmp_newLead) THEN
            tmp_newLead := i;
        END_IF;
    END_FOR;
    leadPump := tmp_newLead;
    tmp_selectLag := TRUE;
    IF demand >= 2 THEN
        newLag := 0;
        FOR i := 1 TO 5 DO
            IF i <> leadPump THEN
                IF newLag = 0 OR runHours[i] < runHours[newLag] OR (runHours[i] = runHours[newLag] AND i < newLag) THEN
                    newLag := i;
                END_IF;
            END_IF;
        END_FOR;
        lagPump := newLag;
    ELSE
        lagPump := 0;
    END_IF;
ELSE
    runningCount := demand;
    IF rotated AND runHours[leadPump] > minHours + 50 THEN
        tmp_newLead := 1;
        FOR i := 2 TO 5 DO
            IF runHours[i] < runHours[tmp_newLead] OR (runHours[i] = runHours[tmp_newLead] AND i < tmp_newLead) THEN
                tmp_newLead := i;
            END_IF;
        END_FOR;
        leadPump := tmp_newLead;
        tmp_selectLag := TRUE;
    END_IF;
    IF demand > tmp_prevRunning THEN
        tmp_newLead := 1;
        FOR i := 2 TO 5 DO
            IF runHours[i] < runHours[tmp_newLead] OR (runHours[i] = runHours[tmp_newLead] AND i < tmp_newLead) THEN
                tmp_newLead := i;
            END_IF;
        END_FOR;
        leadPump := tmp_newLead;
        tmp_selectLag := TRUE;
    END_IF;
    IF tmp_selectLag THEN
        IF demand >= 2 THEN
            newLag := 0;
            FOR i := 1 TO 5 DO
                IF i <> leadPump THEN
                    IF newLag = 0 OR runHours[i] < runHours[newLag] OR (runHours[i] = runHours[newLag] AND i < newLag) THEN
                        newLag := i;
                    END_IF;
                END_IF;
            END_FOR;
            lagPump := newLag;
        ELSE
            lagPump := 0;
        END_IF;
    END_IF;
END_IF;

minHours := runHours[1];
FOR i := 2 TO 5 DO
    IF runHours[i] < minHours THEN
        minHours := runHours[i];
    END_IF;
END_FOR;
END_FUNCTION_BLOCK

(* ---- self-hard-04.raw_candidate_02.st ---- *)
FUNCTION_BLOCK FB
VAR_OUTPUT
    leadPump : INT := 0;
    lagPump : INT := 0;
    runningCount : INT := 0;
END_VAR
VAR_INPUT
    demand : INT;
    runHours : ARRAY[1..5] OF LINT;
    rotated : BOOL;
END_VAR
VAR
    tmp_prevLead : INT := 0;
    tmp_prevRunning : INT := 0;
    tmp_selectLag : BOOL := FALSE;
    tmp_newLead : INT;
    tmp_minOther : LINT;
    i : INT;
END_VAR
VAR_TEMP
    newLag : INT;
    clippedDemand : INT;
END_VAR
(*
ENGINEERING_CONTRACT:
  [S1] runningCount = CLAMP(demand, 0, 5). PUB001/PUB011
  [S2] demand=0→leadPump=lagPump=0; demand=1→lagPump=0; demand≥2→leadPump≠lagPump, both 1..5. PUB002/PUB012
  [S3] Lead-change requires old lead hours > new lead hours + 50. PUB036
  [S4] Hysteresis: rotated=TRUE AND runHours[lead] > minOther + 50 → rotate to min-other pump. PUB026/PUB027
  [S5] Lag pump selected ONLY on: initial, lead change, runningCount increase. PUB005/PUB031
  [S6] Initial lead selection: min (runHours, pump#). PUB028
  [S7] Lag pump: min (runHours, pump#) excluding lead pump. PUB029
  [S8] Demand=0 clears lead/lag immediately; next positive demand triggers fresh selection. PUB033/PUB034
  [S9] First FB invocation initializes all outputs to 0 (VAR_INIT). PUB041
  No edge detection on rotated; it is level-triggered. PUB026
  Array bounds: 1..5 only. PUB042
*)
(* CONTRACT_RULES [] *)

clippedDemand := demand;
IF clippedDemand < 0 THEN
    clippedDemand := 0;
ELSIF clippedDemand > 5 THEN
    clippedDemand := 5;
END_IF;

tmp_prevLead := leadPump;
tmp_prevRunning := runningCount;
tmp_selectLag := FALSE;

IF clippedDemand = 0 THEN
    runningCount := 0;
    leadPump := 0;
    lagPump := 0;
ELSIF leadPump = 0 THEN
    runningCount := clippedDemand;
    tmp_newLead := 1;
    FOR i := 2 TO 5 DO
        IF runHours[i] < runHours[tmp_newLead] OR (runHours[i] = runHours[tmp_newLead] AND i < tmp_newLead) THEN
            tmp_newLead := i;
        END_IF;
    END_FOR;
    leadPump := tmp_newLead;
    tmp_selectLag := TRUE;
    IF clippedDemand >= 2 THEN
        newLag := 0;
        FOR i := 1 TO 5 DO
            IF i <> leadPump THEN
                IF newLag = 0 OR runHours[i] < runHours[newLag] OR (runHours[i] = runHours[newLag] AND i < newLag) THEN
                    newLag := i;
                END_IF;
            END_IF;
        END_FOR;
        lagPump := newLag;
    ELSE
        lagPump := 0;
    END_IF;
ELSE
    runningCount := clippedDemand;
    tmp_minOther := 9223372036854775807; // LINT_MAX approximation
    FOR i := 1 TO 5 DO
        IF i <> leadPump AND runHours[i] < tmp_minOther THEN
            tmp_minOther := runHours[i];
        END_IF;
    END_FOR;
    IF rotated AND runHours[leadPump] > tmp_minOther + 50 THEN
        tmp_newLead := 1;
        FOR i := 2 TO 5 DO
            IF runHours[i] < runHours[tmp_newLead] OR (runHours[i] = runHours[tmp_newLead] AND i < tmp_newLead) THEN
                tmp_newLead := i;
            END_IF;
        END_FOR;
        leadPump := tmp_newLead;
        tmp_selectLag := TRUE;
    END_IF;
    IF clippedDemand > tmp_prevRunning THEN
        tmp_newLead := 1;
        FOR i := 2 TO 5 DO
            IF runHours[i] < runHours[tmp_newLead] OR (runHours[i] = runHours[tmp_newLead] AND i < tmp_newLead) THEN
                tmp_newLead := i;
            END_IF;
        END_FOR;
        leadPump := tmp_newLead;
        tmp_selectLag := TRUE;
    END_IF;
    IF tmp_selectLag THEN
        IF clippedDemand >= 2 THEN
            newLag := 0;
            FOR i := 1 TO 5 DO
                IF i <> leadPump THEN
                    IF newLag = 0 OR runHours[i] < runHours[newLag] OR (runHours[i] = runHours[newLag] AND i < newLag) THEN
                        newLag := i;
                    END_IF;
                END_IF;
            END_FOR;
            lagPump := newLag;
        ELSE
            lagPump := 0;
        END_IF;
    END_IF;
END_IF;
END_FUNCTION_BLOCK

(* ---- self-hard-04.raw_candidate_03.st ---- *)
FUNCTION_BLOCK FB
VAR_OUTPUT
    leadPump : INT := 0;
    lagPump : INT := 0;
    runningCount : INT := 0;
END_VAR
VAR_INPUT
    demand : INT;
    runHours : ARRAY[1..5] OF LINT;
    rotated : BOOL;
END_VAR
VAR
    tmp_prevLead : INT := 0;
    tmp_prevRunning : INT := 0;
    tmp_selectLag : BOOL := FALSE;
    tmp_newLead : INT;
    minHours : LINT;
    i : INT;
    tmp_demand : INT;
END_VAR
VAR_TEMP
    newLag : INT;
END_VAR
(*
ENGINEERING_CONTRACT:
  [S1] runningCount = CLAMP(demand, 0, 5). PUB001/PUB011
  [S2] demand=0→leadPump=lagPump=0; demand=1→lagPump=0; demand≥2→leadPump≠lagPump, both 1..5. PUB002/PUB012
  [S3] Lead-change requires old lead hours > new lead hours + 50. PUB036
  [S4] Hysteresis: rotated=TRUE AND runHours[lead] > minHours + 50 → rotate to min-hours pump. PUB026/PUB027
  [S5] Lag pump selected ONLY on: initial, lead change, runningCount increase. PUB005/PUB031
  [S6] Initial lead selection: min (runHours, pump#). PUB028
  [S7] Lag pump: min (runHours, pump#) excluding lead pump. PUB029
  [S8] Demand=0 clears lead/lag immediately; next positive demand triggers fresh selection. PUB033/PUB034
  [S9] First FB invocation initializes all outputs to 0 (VAR_INIT). PUB041
  No edge detection on rotated; it is level-triggered. PUB026
  Array bounds: 1..5 only. PUB042
*)
(* CONTRACT_RULES [] *)

tmp_prevLead := leadPump;
tmp_prevRunning := runningCount;
tmp_selectLag := FALSE;

IF demand < 0 THEN
    tmp_demand := 0;
ELSIF demand > 5 THEN
    tmp_demand := 5;
ELSE
    tmp_demand := demand;
END_IF;

minHours := runHours[1];
FOR i := 2 TO 5 DO
    IF runHours[i] < minHours THEN
        minHours := runHours[i];
    END_IF;
END_FOR;

IF tmp_demand <= 0 THEN
    runningCount := 0;
    leadPump := 0;
    lagPump := 0;
ELSIF tmp_prevLead = 0 THEN
    runningCount := tmp_demand;
    tmp_newLead := 1;
    FOR i := 2 TO 5 DO
        IF runHours[i] < runHours[tmp_newLead] OR (runHours[i] = runHours[tmp_newLead] AND i < tmp_newLead) THEN
            tmp_newLead := i;
        END_IF;
    END_FOR;
    leadPump := tmp_newLead;
    tmp_selectLag := TRUE;
    IF tmp_demand >= 2 THEN
        newLag := 0;
        FOR i := 1 TO 5 DO
            IF i <> leadPump THEN
                IF newLag = 0 OR runHours[i] < runHours[newLag] OR (runHours[i] = runHours[newLag] AND i < newLag) THEN
                    newLag := i;
                END_IF;
            END_IF;
        END_FOR;
        lagPump := newLag;
    ELSE
        lagPump := 0;
    END_IF;
ELSE
    runningCount := tmp_demand;
    IF rotated AND runHours[leadPump] > minHours + 50 THEN
        tmp_newLead := 1;
        FOR i := 2 TO 5 DO
            IF runHours[i] < runHours[tmp_newLead] OR (runHours[i] = runHours[tmp_newLead] AND i < tmp_newLead) THEN
                tmp_newLead := i;
            END_IF;
        END_FOR;
        leadPump := tmp_newLead;
        tmp_selectLag := TRUE;
    END_IF;
    IF tmp_demand > tmp_prevRunning THEN
        tmp_newLead := 1;
        FOR i := 2 TO 5 DO
            IF runHours[i] < runHours[tmp_newLead] OR (runHours[i] = runHours[tmp_newLead] AND i < tmp_newLead) THEN
                tmp_newLead := i;
            END_IF;
        END_FOR;
        leadPump := tmp_newLead;
        tmp_selectLag := TRUE;
    END_IF;
    IF tmp_selectLag THEN
        IF tmp_demand >= 2 THEN
            newLag := 0;
            FOR i := 1 TO 5 DO
                IF i <> leadPump THEN
                    IF newLag = 0 OR runHours[i] < runHours[newLag] OR (runHours[i] = runHours[newLag] AND i < newLag) THEN
                        newLag := i;
                    END_IF;
                END_IF;
            END_FOR;
            lagPump := newLag;
        ELSE
            lagPump := 0;
        END_IF;
    END_IF;
END_IF;
END_FUNCTION_BLOCK
